// TIA Portal project "Project2" (V17)

(* hardware
DEVICE "S7-1500/ET200MP station_1"  S7-1500 station
   slot 0: "Rail_0"  Rack  6ES7 590-1***0-0AA0
   slot 1: "PLC_2"  CPU 1515-2 PN  6ES7 515-2AM00-0AB0  V1.8
      slot 3: "CPU display_1"  6ES7591-1BA00-0AA0
      slot 32768: "PROFINET interface_1"  X1
         slot 32769: "Port_1"  X1 P1
         slot 32770: "Port_2"  X1 P2
      slot 33024: "PROFINET interface_2"  X2
         slot 33025: "Port_1"  X2 P1
*)

// ===== PLC "PLC_2"  CPU 1515-2 PN =====

// folder: UDT/S2-Process Function Unit

TYPE "UDT_IS28xx_To_Plc"
   STRUCT
      iTriggerReady : Bool;   // This bit indicates when an In-Sight device can accept a new trigger via the Trigger bit. This field is true when the Trigger Enable bit is set, and the vision system is not currently acquiring an image.
      iTriggerAck : Bool;   // This bit indicates when an In-Sight device is successfully triggered via the Trigger bit. The Trigger Acknowledge bit stays set until the Trigger bit is cleared.
      iExposureComplete : Bool;   // This bit is set when the vision system image sensor is no longer exposed to light. It is used to indicate that the part being inspected can be moved from under the vision system's field of view.
      iAcquisitionError : Bool;   // This bit is set when an In-Sight device fails to acquire an image for one of the following reasons:
      iOfflineReason_1 : Bool;   // OfflineReason_1
      iOfflineReason_2 : Bool;   // OfflineReason_2
      iOfflineReason_3 : Bool;   // OfflineReason_3
      iSystemOnline : Bool;   // This bit indicates that the In-Sight device is online and the $System.OnlineEnabled tag is True.
      iReserve_1 : Byte;   // Reserve1
      iAcquisitonID : Int;   // This ID increments on the completion of every acquisition, regardless of the trigger source, and can be used to synchronize an acquisition with its Inspection Result. The Acquisition ID is changed on the start of an acquisition. If the PLC is the trigger source, the Acquisition ID is set prior to setting the Trigger Acknowledge bit.
      iReserve_2 : Bool;   // Reserve2
      iInspectionComplete : Bool;   // This bit is toggled upon the completion of an inspection.
      iResultBufferOverRun : Bool;   // This bit is set when the Enable Results Buffer bit is set, and there are more results than the result queue can hold.
      iResultValid : Bool;   // This bit is set when the Inspected Image ID, Inspection Result Code and Inspection Results fields are valid. The bit is cleared when the Inspection Results Acknowledge bit is set.
      iCommandExecuted : Bool;   // This bit is set while a command execution is in progress.
      iCommandComplete : Bool;   // This bit is set when the command execution is completed, and cleared when the Execute Command bit has been cleare
      iCommandFailed : Bool;   // This bit is set on the completion of a command, if the command has failed to execute successfully, or if an unknown Command ID was set.
      iSetUserDataAck : Bool;   // This bit is set to acknowledge completion of the Set User Data command.
      iJobPass : Bool;   // This bit indicates the pass and/or fail state of the inspection.
      iReserve_3 : Bool;   // Reserve3
      iReserve_4 : Bool;   // Reserve4
      iReserve_5 : Bool;   // Reserve5
      iReserve_6 : Bool;   // Reserve6
      iReserve_7 : Bool;   // Reserve7
      iReserve_8 : Bool;   // Reserve8
      iError : Bool;   // This bit is set when an error has occurred, which is defined in the Error ID field.
      iErrorID : Int;   // See Error ID codes.
      iCurrentRunningJobID : Int;   // These bits indicate the pre-added number of the current job filename. A job ID is a 16 bit number from 0 to 65535, but the PLC function can only load job IDs between 0‑999.
      iCommandResultCode : Int;   // This field is used to indicate the reason a command failed to execute successfully (the code is specific to the command executed):
      iExternalSoftEventAck : Byte;   // The External Event Acknowledge will be generated after the associated script finishes its execution
      iInspectionResultData : Struct
         iInspectionID : Int;   // The acquisition ID associated with this set of results.
         iInspectionResultCode : Int;   // These bytes are used to pass the user-defined result code. The inspection result code is defined by the Result Code parameter of the WriteResultsBuffer function
         iInspectionResult : Array[1..60] of Byte;   // These bytes of the inspection tool results can be written to the currently enabled factory communication protocol via the WriteResultsBuffer function.
      END_STRUCT;
   END_STRUCT;
END_TYPE

TYPE "UDT_Plc_To_IS28xx"
   STRUCT
      qTriggerEnable : Bool;   // This field is set to enable triggering via the Trigger bit. Clear this bit to disable the network triggering mechanism
      qTrigger : Bool;   // Setting the Trigger bit will trigger an acquisition on the vision system. The Trigger Enable bit must also be set
      qClearExposureComplete : Bool;   // When this signal is held high, the Exposure Complete status will remain reset. Once this signal is set to low, the Exposure Complete status will be set to high on the next exposure completion.
      qReserve_1 : Bool;   // Reserve_1
      qReserve_2 : Bool;   // Reserve_2
      qReserve_3 : Bool;   // Reserve_3
      qReserve_4 : Bool;   // Reserve_4
      qSetOffline : Bool;   // When this bit is set, the In-Sight vision system is paused and the state of the $System.OnlineEnabledComm is false
      qBufferResultEnable : Bool;   // When this bit is set, the Inspection ID, Inspection Result and Inspection Results fields are held constant until the Inspection Results Acknowledge field has acknowledged them and been set. Up to 16 sets of results are held in the buffer. Each result must be explicitly acknowledged using the Inspection Results Acknowledge signal.
      qInspectionResultAck : Bool;   // When the Buffer Results Enable bit is set, the Inspection Results Acknowledge bit acknowledges that the PLC has received the Inspected Image ID, Inspection Result Code and Inspection Results data.
      qSetUserData : Bool;   // This bit is used to signal that new User Data is available to be read in the vision system. After latching the entire User Data area into a holding buffer, the vision system will indicate to the PLC that it has read the data, and it can start loading new data into the buffer, if required, by issuing the Set User Data Acknowledge signal.
      qExecuteCommand : Bool;   // When the Execute Command bit is set to high, the Command ID signal is read by the vision system and the associated command is executed. The signal must be held high until the Command Completed bit is set. Once the Command Completed bit is set, clearing the Execute Command bit also clears the Command Completed bit.
      qReserve_5 : Bool;   // Reserve_5
      qReserve_6 : Bool;   // Reserve_6
      qReserve_7 : Bool;   // Reserve_7
      qClearError : Bool;   // When this bit is set, it clears the Error and Error ID signals; the Clear Error bit need to be held high until the Error bit is cleared. If an error is queued, clearing this bit causes the Error and Error ID signals to be set to the next queued error code.
      qCommandID : Int;   // This field indicates the command that will be executed on the rising edge of the Execute Command bit. This signal should not be changed until the Command Completed bit has been set.
      qSoftControlInput : Byte;   // Setting the External Event allows the PLC to trigger an associated event in the Spreadsheet.
      qUserData : Array[1..60] of Byte;   // Data buffer which can be read into the spreadsheet using the ReadUserDataBuffer function. The buffer is written exactly as it appears in the PLC
   END_STRUCT;
END_TYPE

// folder: (top level)

ORGANIZATION_BLOCK "Main"   // OB1, LAD, ProgramCycle
TITLE = "Main Program Sweep (Cycle)"
{ S7_Optimized_Access := 'TRUE' }
VERSION : 0.1
   VAR_INPUT
      Initial_Call : Bool;   // Initial call of this OB
      Remanence : Bool;   // =True, if remanent data are available
   END_VAR
   VAR_TEMP
      OB1_EV_CLASS : Byte;   // Bits 0-3 = 1 (Coming event), Bits 4-7 = 1 (Event class 1)
      OB1_SCAN_1 : Byte;   // 1 (Cold restart scan 1 of OB 1), 3 (Scan 2-n of OB 1)
      OB1_PRIORITY : Byte;   // Priority of OB Execution
      OB1_OB_NUMBR : Byte;   // 1 (Organization block 1, OB1)
      OB1_RESERVED_1 : Byte;   // Reserved for system
      OB1_RESERVED_2 : Byte;   // Reserved for system
      OB1_PREV_CYCLE : Int;   // Cycle time of previous OB1 scan (milliseconds)
      OB1_MIN_CYCLE : Int;   // Minimum cycle time of OB1 (milliseconds)
      OB1_MAX_CYCLE : Int;   // Maximum cycle time of OB1 (milliseconds)
      OB1_DATE_TIME : Date_And_Time;   // Date and time OB1 started
   END_VAR
BEGIN
END_ORGANIZATION_BLOCK

// ===== library types =====

// folder: S2-Process Function Unit

FUNCTION_BLOCK "PR_CognexISCamera_Profinet"   // FB365, LAD
TITLE = Cognex2D_4Feature / Cognex Camera Module
{ S7_Optimized_Access := 'TRUE' }
AUTHOR : Deepak.Jagtap
FAMILY : WIPROPARI
NAME : S21006022005
VERSION : 0.1
// |============================================================================|
// BLOCK:Cognex Camera Module
// Item Code : SMxxxxx
// Owner:Precision Automation & Robotics India Ltd.
// Author: DJ
// Release Date:04-04-2018
// Version:0.1
// V0.1-Initial release
// |============================================================================|
// Block Description: This block is used for interface of Cognex Camera via 
// profinet  and enter Job selection from outside the block.
// |============================================================================|
// Errors:
// qErrTriggerTimeOut: Trigger TimeOut Error Occured
// qErrAcquiringTimeout: Acquiring TimeOut Error Occured
// qErrTriggerEnableTimeout: Trigger Enable TimeOut Occured
// qErrJobSelection: Job selection Error
// qBothStartOn: Both Start are ON
// ============================================================================|
// Dependency:
// Map Vision Input and Output from External IO address. Byte should be matched as per the block
// |============================================================================|
   VAR_INPUT
      iResetFault : Bool;   // Reset Fault Input
      iAutorunning : Bool;   // Autorunning Input
      iStartJobSelection : Bool;   // start job selection / Start for Job Selection
      iStartInspection : Bool;   // Start for Inspection / start inspection
      iRetryCount : Int;   // Retry Count eg:3,4 etc / retry count
      iRetryPB : Bool;
      iJobID : Int;   // Enter Job ID / job id
      iTriggerEnableTimeoutTime : Time;   // Trigger Enable TimeOut Time Delay
      iTriggerTimeoutTime : Time;   // Trigger TimeOut Time Delay
      iAcquiringTimeOutTime : Time;   // Acquiring TimeOut Time Delay
   END_VAR
   VAR_OUTPUT
      qJobPass : Bool;   // Job Pass In Inspection
      qJobFail : Bool;   // Job Failed In Inspection
      qJobSelectionOver : Bool;   // Connect Job Selection over bit / job selection over
      qJobInspectionOver : Bool;   // Inspection Over Output
      qVisionOnline : Bool;   // Insight Vision Is In Online
      qVisionOfflineReason1 : Bool;   // Insight Vision Offline Due To: The vision system's job is being modified
      qVisionOfflineReason2 : Bool;   // Insight Vision Offline Due To: A discrete signal is holding the vision system Offline
      qVisionOfflineReason3 : Bool;   // Insight Vision Offline Due To: A communications protocol is holding the vision system Offline
      qErrBothStartOn : Bool;   // Both Start are On / both start on
      qErrJobSelection : Bool;   // Job selection Error Occur / error job selection
      qErrTriggerEnableTimeout : Bool;   // Trigger Enable TimeOut Error
      qErrTriggerTimeOut : Bool;   // Trigger TimeOut Error
      qErrAcquiringTimeOut : Bool;   // Acquiring TimeOut Error
   END_VAR
   VAR_IN_OUT
      iqInputAddrs : ANY;   // Input HW Address P#I120.0 BYTE 74
      iqOutputAddrs : ANY;   // Input HW Address P#Q120.0 BYTE 68
      iqRetryCount : Int;   // Retry Count Display / Retry count
      iqRunningJobID : Int;   // Running job ID
      iqInsight_Camera : Struct   // Insight Camera PZD
         Vision_Input : Struct
            "iTrigger Ready" : Bool;
            "iTrigger Ack" : Bool;
            iExposureComplete : Bool;
            "iMissed Ack" : Bool;
            "iOffline Reason_0" : Bool;
            "iOffline Reason_1" : Bool;
            "iOffline Reason_2" : Bool;
            iOnline : Bool;
            Acquisition_ID : Byte;
            Acquisition_ID_1 : Byte;
            iSystemBusy : Bool;
            "iInspection Completed" : Bool;
            "iResults Buffer Overrun" : Bool;
            "iResults Valid" : Bool;
            iCommandExecuting : Bool;
            iCommandComplete : Bool;
            "iCommand Failed" : Bool;
            iSetUserDataAck : Bool;
            iJobPass : Bool;
            iReserved : Bool;
            iReserved_1 : Bool;
            iReserved_2 : Bool;
            iReserved_3 : Bool;
            iReserved_4 : Bool;
            iReserved_5 : Bool;
            iError : Bool;
            iErrorCode : Int;
            iCommandControlInput : Int;
            SoftEventControlInput : Byte;
            iInspection_ID : Byte;
            iInspection_ID_1 : Byte;
            iInspection_ResultCode : Byte;
            iInspection_ResultCode_1 : Byte;
            iInspection_Result : Array[213..277] of Byte;
         END_STRUCT;
         Vision_Output : Struct
            "qTrigger Enable" : Bool;
            qTrigger : Bool;
            qClearExposureComplete : Bool;
            qReserved_1 : Bool;
            qReserved_2 : Bool;
            qReserved_3 : Bool;
            qReserved_4 : Bool;
            "qSet Offline" : Bool;
            "qBuffer Results Enable" : Bool;
            "qInspection Results Ack" : Bool;
            qSetUserData : Bool;
            qExecuteCommand : Bool;
            qReserved : Bool;
            qReserved_5 : Bool;
            qReserved_6 : Bool;
            qClearError : Bool;
            qCommandControl : Word;
            "Soft Event Control" : Byte;
            qUser_Data : Array[205..268] of Byte;
         END_STRUCT;
      END_STRUCT;
   END_VAR
   VAR
      sResetFaults : Bool;   // Reset Faults
      sInspectionComplete : Bool;   // Inspection Complete
      TriggerTimeout : TON_TIME;   // TriggerTimeout Timer
      TriggerEnableTimeout : TON_TIME;   // TriggerEnableTimeout Timer
      AcquiringTimeOut : TON_TIME;   // AcquiringTimeOut Timer
      ResultTimer : TON_TIME;   // ResultTimer
      sPulse : Array[0..11] of Bool;   // Array of Pulses
      sJobPass : Bool;   // Stat Bit of Job Pass
      sVisionInputCmdControlIP : Int;
      sJobFail : Bool;   // Stat Bit of Job Fail
      sJobLoadcompleted : Bool;
      sErrTriggerTimeOut : Bool;   // Error Trigger Time Out
      sErrJobSelection : Bool;
      sBothStartOn : Bool;
      sJobSelectionOver : Bool;
      sJobInspectionOver : Bool;
      sErrAcquiringTimeOut : Bool;   // Error Acquiring Time Out
      sErrTriggerEnableTimeout : Bool;   // Error Trigger Enable Time Out
      sVisionOutput_Trigger : Bool;   // Vision Outpur Trigger
      sRetryCountOver : Bool;
      sInitialPulse : Bool;
      sProgramEcho : TON_TIME;
      sExposureTimerStar1 : Bool;
      sExposureTimerStart : Bool;
      sExposureTimer : TON_TIME;
      sExecDelayTimer : TON_TIME;
      sRetry : TON_TIME;
   END_VAR
   VAR_TEMP
      tInspectionID : Int;
      tResultCode : Int;
   END_VAR
   VAR_TEMP   // added for the SCL form of the ladder/FBD networks
      _w1 : Bool;
      _w2 : Bool;
      _w3 : Bool;
      _w4 : Bool;
   END_VAR
BEGIN

REGION Network 1: Header
   // ==============================================================================
   //  Company: Precision Automation & Robotics India Ltd. 
   // ------------------------------------------------------------------------------
   //  Item Code: S21006022005
   //  Author/Created by: Deepak.Jagtap
   //  Reviewed/Checked by: Atul P
   //  First Release on: 04-04-2018
   //  Latest update on:
   // ------------------------------------------------------------------------------
   //  Tested with: CPU firmware, model or simulator testing
   //  Engineering/Editor: TIA Portal V15.1
   // ------------------------------------------------------------------------------
   //  Restrictions:
   //  Dependencies/Requirements:
   // iqInsight_Camera	Struct
   // Map Vision Input and Output from with External IO address
   // ------------------------------------------------------------------------------
   //  Change Log:
   //  Ver.	Date		Changed by		Details of changes
   //  1.0	04-04-2018	Deepak.Jagtap            	First release version
   // 
   // ------------------------------------------------------------------------------
   //  Functionality: This block is used for interface of Cognex Camera via 
   // profinet.
   // 
   //  Inputs
   // iResetFault	Bool
   // iAutorunning	Bool
   // iStartJobSelection	Bool
   // iStartInspection	Bool
   // iRetryCount	Int
   // iJobID	Int
   // iTriggerEnableTimeoutTime	Time
   // iTriggerTimeoutTime	Time
   // iAcquiringTimeOutTime	Time
   // 
   //  Outputs
   // qJobPass	Bool
   // qJobFail	Bool
   // qJobSelectionOver	Bool
   // qJobInspectionOver	Bool
   // qVisionOnline	Bool
   // qVisionOfflineReason1	Bool
   // qVisionOfflineReason2	Bool
   // qVisionOfflineReason3	Bool
   // qErrBothStartOn	Bool
   // qErrJobSelection	Bool
   // qErrTriggerEnableTimeout	Bool
   // qErrTriggerTimeOut	Bool
   // qErrAcquiringTimeOut	Bool
   // 
   //  In-outs
   // iqInputAddrs	Any
   // iqOutputAddrs	Any
   // iqRetryCount	Int
   // iqRunningJobID	Int
   // iqInsight_Camera	Struct
   // 
   // ------------------------------------------------------------------------------
   //  Errors reported:
   //  1.qErrTriggerTimeOut : Error trigger timeout
   // 2. qErrAcquiringTimeOut;Acquiring Time Out
   // 3. qErrTriggerEnableTimeout:Trigger Enable Time Out
   // 4. qErrBothStartOn:both start on
   // 5. qErrJobSelection:error job selection
   //  Messages reported:
   //  1. Message 1 present
   //  2. Message 2 present
   // ==============================================================================
END_REGION

REGION Network 2: Read Data From Input Area
   // Read Data From Input Area
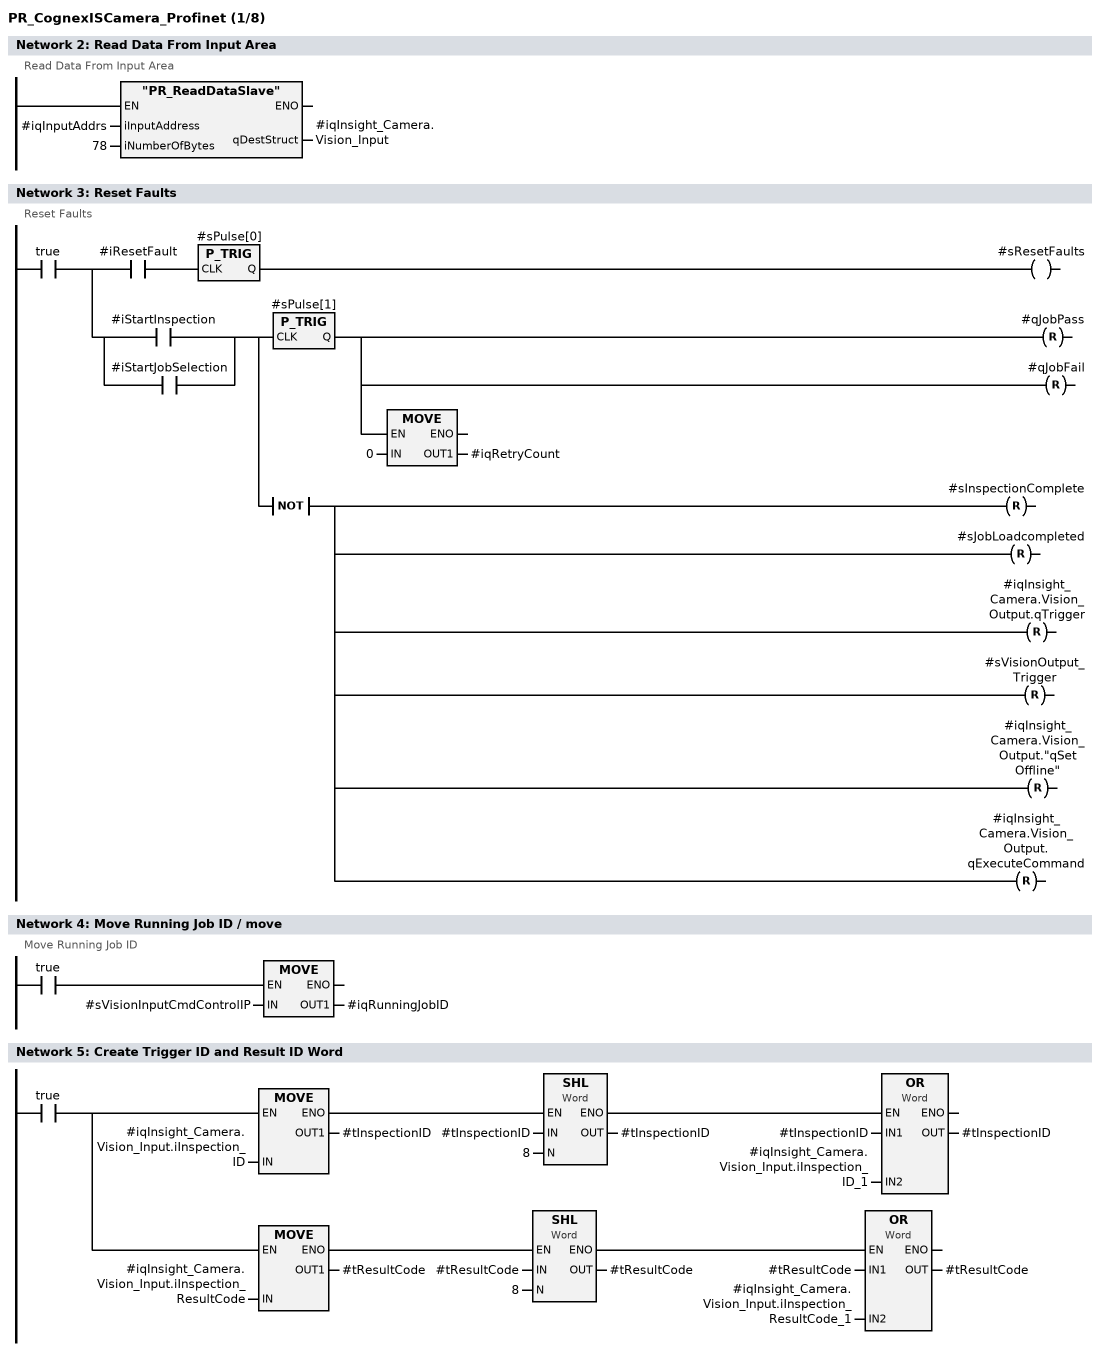
   RUNG wire#powerrail
      "PR_ReadDataSlave"(iInputAddress := #iqInputAddrs, iNumberOfBytes := 78, qDestStruct => #iqInsight_Camera.Vision_Input)
   END_RUNG
   // the same network as SCL:
   "PR_ReadDataSlave"(iInputAddress := #iqInputAddrs,
                      iNumberOfBytes := 78,
                      qDestStruct => #iqInsight_Camera.Vision_Input);
END_REGION

REGION Network 3: Reset Faults
   // Reset Faults
   RUNG wire#powerrail
      Contact( true )
      wire#w1
      Contact( #iResetFault )
      P_Trig( #sPulse[0] )
      Coil( #sResetFaults )
   END_RUNG
   RUNG wire#w1
      Contact( #iStartInspection )
      wire#w2
      P_Trig( #sPulse[1] )
      wire#w3
      R_Coil( #qJobPass )
   END_RUNG
   RUNG wire#w1
      Contact( #iStartJobSelection )
   END_RUNG wire#w2
   RUNG wire#w3
      R_Coil( #qJobFail )
   END_RUNG
   RUNG wire#w3
      Move(in := 0, out1 => #iqRetryCount)
   END_RUNG
   RUNG wire#w2
      Not()
      wire#w4
      R_Coil( #sInspectionComplete )
   END_RUNG
   RUNG wire#w4
      R_Coil( #sJobLoadcompleted )
   END_RUNG
   RUNG wire#w4
      R_Coil( #iqInsight_Camera.Vision_Output.qTrigger )
   END_RUNG
   RUNG wire#w4
      R_Coil( #sVisionOutput_Trigger )
   END_RUNG
   RUNG wire#w4
      R_Coil( #iqInsight_Camera.Vision_Output."qSet Offline" )
   END_RUNG
   RUNG wire#w4
      R_Coil( #iqInsight_Camera.Vision_Output.qExecuteCommand )
   END_RUNG
   // the same network as SCL:
   #_w1 := true AND #iResetFault;
   #_w2 := #_w1 AND NOT #sPulse[0];   // rising edge
   #sPulse[0] := #_w1;
   #sResetFaults := #_w2;
   #_w3 := true AND (#iStartInspection OR #iStartJobSelection);
   #_w4 := #_w3 AND NOT #sPulse[1];   // rising edge
   #sPulse[1] := #_w3;
   IF #_w4 THEN
       #qJobPass := FALSE;
       #qJobFail := FALSE;
       #iqRetryCount := 0;
   END_IF;
   IF NOT #_w3 THEN
       #sInspectionComplete := FALSE;
       #sJobLoadcompleted := FALSE;
       #iqInsight_Camera.Vision_Output.qTrigger := FALSE;
       #sVisionOutput_Trigger := FALSE;
       #iqInsight_Camera.Vision_Output."qSet Offline" := FALSE;
       #iqInsight_Camera.Vision_Output.qExecuteCommand := FALSE;
   END_IF;
END_REGION

REGION Network 4: Move Running Job ID / move
   // Move Running Job ID
   RUNG wire#powerrail
      Contact( true )
      Move(in := #sVisionInputCmdControlIP, out1 => #iqRunningJobID)
   END_RUNG
   // the same network as SCL:
   IF true THEN #iqRunningJobID := #sVisionInputCmdControlIP; END_IF;
END_REGION

REGION Network 5: Create Trigger ID and Result ID Word
   IF true THEN
       #tInspectionID := #iqInsight_Camera.Vision_Input.iInspection_ID;
       #tInspectionID := SHL(IN := #tInspectionID, N := 8);
       #tInspectionID := #tInspectionID OR #iqInsight_Camera.Vision_Input.iInspection_ID_1;
       #tResultCode := #iqInsight_Camera.Vision_Input.iInspection_ResultCode;
       #tResultCode := SHL(IN := #tResultCode, N := 8);
       #tResultCode := #tResultCode OR #iqInsight_Camera.Vision_Input.iInspection_ResultCode_1;
   END_IF;
END_REGION

REGION Network 6: Trigger Enable through Job Selection / Camera Trigger Enable
   // Trigger Enable through Job Selection
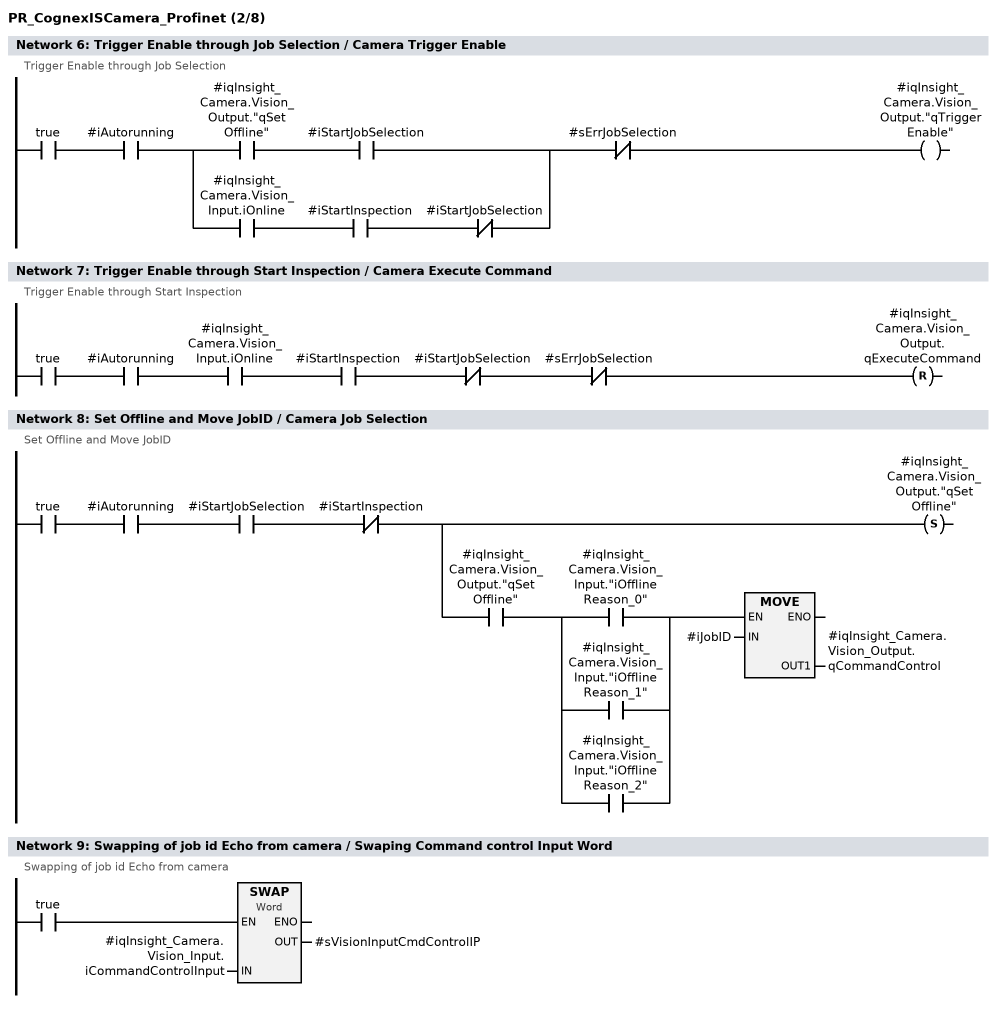
   RUNG wire#powerrail
      Contact( true )
      Contact( #iAutorunning )
      wire#w1
      Contact( #iqInsight_Camera.Vision_Output."qSet Offline" )
      Contact( #iStartJobSelection )
      wire#w2
      I_Contact( #sErrJobSelection )
      Coil( #iqInsight_Camera.Vision_Output."qTrigger Enable" )
   END_RUNG
   RUNG wire#w1
      Contact( #iqInsight_Camera.Vision_Input.iOnline )
      Contact( #iStartInspection )
      I_Contact( #iStartJobSelection )
   END_RUNG wire#w2
   // the same network as SCL:
   #iqInsight_Camera.Vision_Output."qTrigger Enable" := true AND #iAutorunning AND ((#iqInsight_Camera.Vision_Output."qSet Offline" AND #iStartJobSelection) OR (#iqInsight_Camera.Vision_Input.iOnline AND #iStartInspection AND NOT #iStartJobSelection)) AND NOT #sErrJobSelection;
END_REGION

REGION Network 7: Trigger Enable through Start Inspection / Camera Execute Command
   // Trigger Enable through Start Inspection
   RUNG wire#powerrail
      Contact( true )
      Contact( #iAutorunning )
      Contact( #iqInsight_Camera.Vision_Input.iOnline )
      Contact( #iStartInspection )
      I_Contact( #iStartJobSelection )
      I_Contact( #sErrJobSelection )
      R_Coil( #iqInsight_Camera.Vision_Output.qExecuteCommand )
   END_RUNG
   // the same network as SCL:
   IF true AND #iAutorunning AND #iqInsight_Camera.Vision_Input.iOnline AND #iStartInspection AND NOT #iStartJobSelection AND NOT #sErrJobSelection THEN
       #iqInsight_Camera.Vision_Output.qExecuteCommand := FALSE;
   END_IF;
END_REGION

REGION Network 8: Set Offline and Move JobID / Camera Job Selection
   // Set Offline and Move JobID
   RUNG wire#powerrail
      Contact( true )
      Contact( #iAutorunning )
      Contact( #iStartJobSelection )
      I_Contact( #iStartInspection )
      wire#w1
      S_Coil( #iqInsight_Camera.Vision_Output."qSet Offline" )
   END_RUNG
   RUNG wire#w1
      Contact( #iqInsight_Camera.Vision_Output."qSet Offline" )
      wire#w2
      Contact( #iqInsight_Camera.Vision_Input."iOffline Reason_0" )
      wire#w3
      Move(in := #iJobID, out1 => #iqInsight_Camera.Vision_Output.qCommandControl)
   END_RUNG
   RUNG wire#w2
      Contact( #iqInsight_Camera.Vision_Input."iOffline Reason_1" )
   END_RUNG wire#w3
   RUNG wire#w2
      Contact( #iqInsight_Camera.Vision_Input."iOffline Reason_2" )
   END_RUNG wire#w3
   // the same network as SCL:
   #_w1 := true AND #iAutorunning AND #iStartJobSelection AND NOT #iStartInspection;
   IF #_w1 THEN #iqInsight_Camera.Vision_Output."qSet Offline" := TRUE; END_IF;
   IF #_w1 AND #iqInsight_Camera.Vision_Output."qSet Offline" AND (#iqInsight_Camera.Vision_Input."iOffline Reason_0" OR #iqInsight_Camera.Vision_Input."iOffline Reason_1" OR #iqInsight_Camera.Vision_Input."iOffline Reason_2") THEN
       #iqInsight_Camera.Vision_Output.qCommandControl := #iJobID;
   END_IF;
END_REGION

REGION Network 9: Swapping of job id Echo from camera / Swaping Command control Input Word
   // Swapping of job id Echo from camera
   IF true THEN
       #sVisionInputCmdControlIP := SWAP(#iqInsight_Camera.Vision_Input.iCommandControlInput);
   END_IF;
END_REGION

REGION Network 10: Initiate Job Load / Camera Execute Command
   // Initiate Job Load
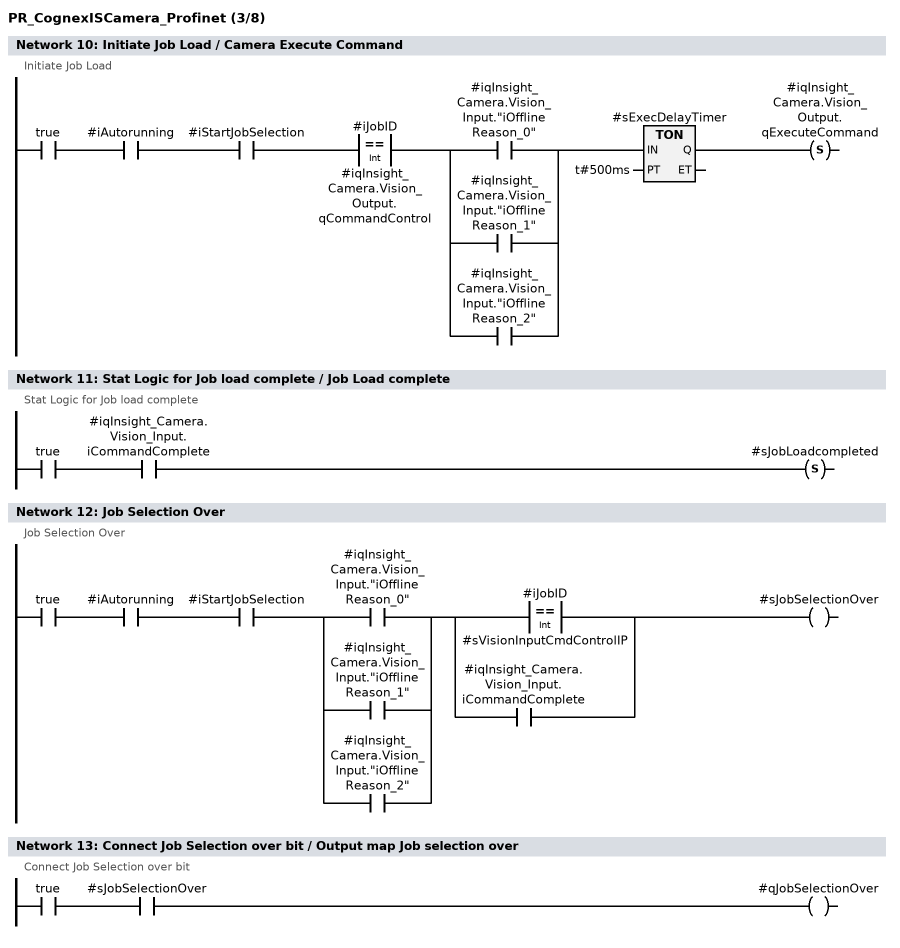
   #sExecDelayTimer(IN := true AND #iAutorunning AND #iStartJobSelection AND (#iJobID = #iqInsight_Camera.Vision_Output.qCommandControl) AND (#iqInsight_Camera.Vision_Input."iOffline Reason_0" OR #iqInsight_Camera.Vision_Input."iOffline Reason_1" OR #iqInsight_Camera.Vision_Input."iOffline Reason_2"),   // TON
                    PT := t#500ms);
   IF #sExecDelayTimer.Q THEN #iqInsight_Camera.Vision_Output.qExecuteCommand := TRUE; END_IF;
END_REGION

REGION Network 11: Stat Logic for Job load complete / Job Load complete
   // Stat Logic for Job load complete
   RUNG wire#powerrail
      Contact( true )
      Contact( #iqInsight_Camera.Vision_Input.iCommandComplete )
      S_Coil( #sJobLoadcompleted )
   END_RUNG
   // the same network as SCL:
   IF true AND #iqInsight_Camera.Vision_Input.iCommandComplete THEN #sJobLoadcompleted := TRUE; END_IF;
END_REGION

REGION Network 12: Job Selection Over
   // Job Selection Over
   RUNG wire#powerrail
      Contact( true )
      Contact( #iAutorunning )
      Contact( #iStartJobSelection )
      wire#w1
      Contact( #iqInsight_Camera.Vision_Input."iOffline Reason_0" )
      wire#w2
      { S7_Templates := "SrcType := Int" } EQ_Contact(in1 := #iJobID, in2 := #sVisionInputCmdControlIP)
      wire#w3
      Coil( #sJobSelectionOver )
   END_RUNG
   RUNG wire#w1
      Contact( #iqInsight_Camera.Vision_Input."iOffline Reason_1" )
   END_RUNG wire#w2
   RUNG wire#w1
      Contact( #iqInsight_Camera.Vision_Input."iOffline Reason_2" )
   END_RUNG wire#w2
   RUNG wire#w2
      Contact( #iqInsight_Camera.Vision_Input.iCommandComplete )
   END_RUNG wire#w3
   // the same network as SCL:
   #sJobSelectionOver := true AND #iAutorunning AND #iStartJobSelection AND (#iqInsight_Camera.Vision_Input."iOffline Reason_0" OR #iqInsight_Camera.Vision_Input."iOffline Reason_1" OR #iqInsight_Camera.Vision_Input."iOffline Reason_2") AND ((#iJobID = #sVisionInputCmdControlIP) OR #iqInsight_Camera.Vision_Input.iCommandComplete);
END_REGION

REGION Network 13: Connect Job Selection over bit / Output map Job selection over
   // Connect Job Selection over bit
   RUNG wire#powerrail
      Contact( true )
      Contact( #sJobSelectionOver )
      Coil( #qJobSelectionOver )
   END_RUNG
   // the same network as SCL:
   #qJobSelectionOver := true AND #sJobSelectionOver;
END_REGION

REGION Network 14: Reset Offline / Camera Job Selection reset
   // Reset Offline / "#iqInsight_Camera.Vision_Output.qSet Offline" and "#iqInsight_Camera.Vision_Output.qExecuteCommand"  Reset coil removed while block comparision
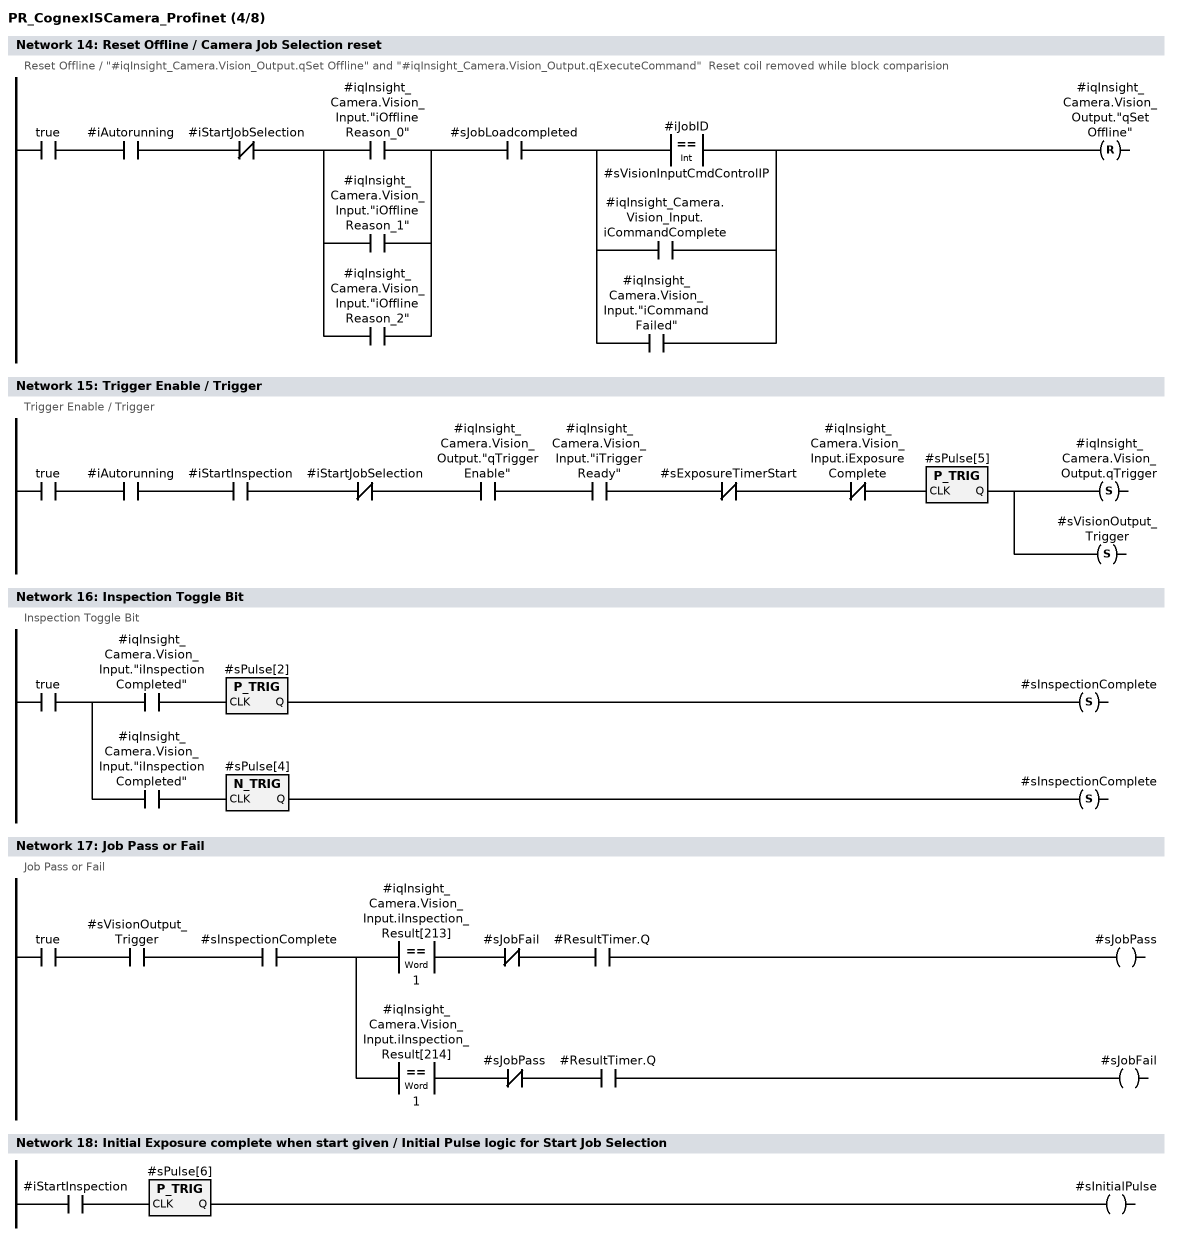
   RUNG wire#powerrail
      Contact( true )
      Contact( #iAutorunning )
      I_Contact( #iStartJobSelection )
      wire#w1
      Contact( #iqInsight_Camera.Vision_Input."iOffline Reason_0" )
      wire#w2
      Contact( #sJobLoadcompleted )
      wire#w3
      { S7_Templates := "SrcType := Int" } EQ_Contact(in1 := #iJobID, in2 := #sVisionInputCmdControlIP)
      wire#w4
      R_Coil( #iqInsight_Camera.Vision_Output."qSet Offline" )
   END_RUNG
   RUNG wire#w1
      Contact( #iqInsight_Camera.Vision_Input."iOffline Reason_1" )
   END_RUNG wire#w2
   RUNG wire#w1
      Contact( #iqInsight_Camera.Vision_Input."iOffline Reason_2" )
   END_RUNG wire#w2
   RUNG wire#w3
      Contact( #iqInsight_Camera.Vision_Input.iCommandComplete )
   END_RUNG wire#w4
   RUNG wire#w3
      Contact( #iqInsight_Camera.Vision_Input."iCommand Failed" )
   END_RUNG wire#w4
   // the same network as SCL:
   IF true AND #iAutorunning AND NOT #iStartJobSelection AND (#iqInsight_Camera.Vision_Input."iOffline Reason_0" OR #iqInsight_Camera.Vision_Input."iOffline Reason_1" OR #iqInsight_Camera.Vision_Input."iOffline Reason_2") AND #sJobLoadcompleted AND ((#iJobID = #sVisionInputCmdControlIP) OR #iqInsight_Camera.Vision_Input.iCommandComplete OR #iqInsight_Camera.Vision_Input."iCommand Failed") THEN
       #iqInsight_Camera.Vision_Output."qSet Offline" := FALSE;
   END_IF;
END_REGION

REGION Network 15: Trigger Enable / Trigger
   // Trigger Enable / Trigger
   RUNG wire#powerrail
      Contact( true )
      Contact( #iAutorunning )
      Contact( #iStartInspection )
      I_Contact( #iStartJobSelection )
      Contact( #iqInsight_Camera.Vision_Output."qTrigger Enable" )
      Contact( #iqInsight_Camera.Vision_Input."iTrigger Ready" )
      I_Contact( #sExposureTimerStart )
      I_Contact( #iqInsight_Camera.Vision_Input.iExposureComplete )
      P_Trig( #sPulse[5] )
      wire#w1
      S_Coil( #iqInsight_Camera.Vision_Output.qTrigger )
   END_RUNG
   RUNG wire#w1
      S_Coil( #sVisionOutput_Trigger )
   END_RUNG
   // the same network as SCL:
   #_w1 := true AND #iAutorunning AND #iStartInspection AND NOT #iStartJobSelection AND #iqInsight_Camera.Vision_Output."qTrigger Enable" AND #iqInsight_Camera.Vision_Input."iTrigger Ready" AND NOT #sExposureTimerStart AND NOT #iqInsight_Camera.Vision_Input.iExposureComplete;
   #_w2 := #_w1 AND NOT #sPulse[5];   // rising edge
   #sPulse[5] := #_w1;
   IF #_w2 THEN
       #iqInsight_Camera.Vision_Output.qTrigger := TRUE;
       #sVisionOutput_Trigger := TRUE;
   END_IF;
END_REGION

REGION Network 16: Inspection Toggle Bit
   // Inspection Toggle Bit
   RUNG wire#powerrail
      Contact( true )
      wire#w1
      Contact( #iqInsight_Camera.Vision_Input."iInspection Completed" )
      P_Trig( #sPulse[2] )
      S_Coil( #sInspectionComplete )
   END_RUNG
   RUNG wire#w1
      Contact( #iqInsight_Camera.Vision_Input."iInspection Completed" )
      N_Trig( #sPulse[4] )
      S_Coil( #sInspectionComplete )
   END_RUNG
   // the same network as SCL:
   #_w1 := true AND #iqInsight_Camera.Vision_Input."iInspection Completed";
   #_w2 := #_w1 AND NOT #sPulse[2];   // rising edge
   #sPulse[2] := #_w1;
   IF #_w2 THEN #sInspectionComplete := TRUE; END_IF;
   #_w3 := true AND #iqInsight_Camera.Vision_Input."iInspection Completed";
   #_w4 := NOT #_w3 AND #sPulse[4];   // falling edge
   #sPulse[4] := #_w3;
   IF #_w4 THEN #sInspectionComplete := TRUE; END_IF;
END_REGION

REGION Network 17: Job Pass or Fail
   // Job Pass or Fail
   RUNG wire#powerrail
      Contact( true )
      Contact( #sVisionOutput_Trigger )
      Contact( #sInspectionComplete )
      wire#w1
      { S7_Templates := "SrcType := Word" } EQ_Contact(in1 := #iqInsight_Camera.Vision_Input.iInspection_Result[213], in2 := 1)
      I_Contact( #sJobFail )
      Contact( #ResultTimer.Q )
      Coil( #sJobPass )
   END_RUNG
   RUNG wire#w1
      { S7_Templates := "SrcType := Word" } EQ_Contact(in1 := #iqInsight_Camera.Vision_Input.iInspection_Result[214], in2 := 1)
      I_Contact( #sJobPass )
      Contact( #ResultTimer.Q )
      Coil( #sJobFail )
   END_RUNG
   // the same network as SCL:
   #_w1 := true AND #sVisionOutput_Trigger AND #sInspectionComplete;
   #sJobPass := #_w1 AND (#iqInsight_Camera.Vision_Input.iInspection_Result[213] = 1) AND NOT #sJobFail AND #ResultTimer.Q;
   #sJobFail := #_w1 AND (#iqInsight_Camera.Vision_Input.iInspection_Result[214] = 1) AND NOT #sJobPass AND #ResultTimer.Q;
END_REGION

REGION Network 18: Initial Exposure complete when start given / Initial Pulse logic for Start Job Selection
   RUNG wire#powerrail
      Contact( #iStartInspection )
      P_Trig( #sPulse[6] )
      Coil( #sInitialPulse )
   END_RUNG
   // the same network as SCL:
   #_w1 := #iStartInspection AND NOT #sPulse[6];   // rising edge
   #sPulse[6] := #iStartInspection;
   #sInitialPulse := #_w1;
END_REGION

REGION Network 19: Exposure Timer 1
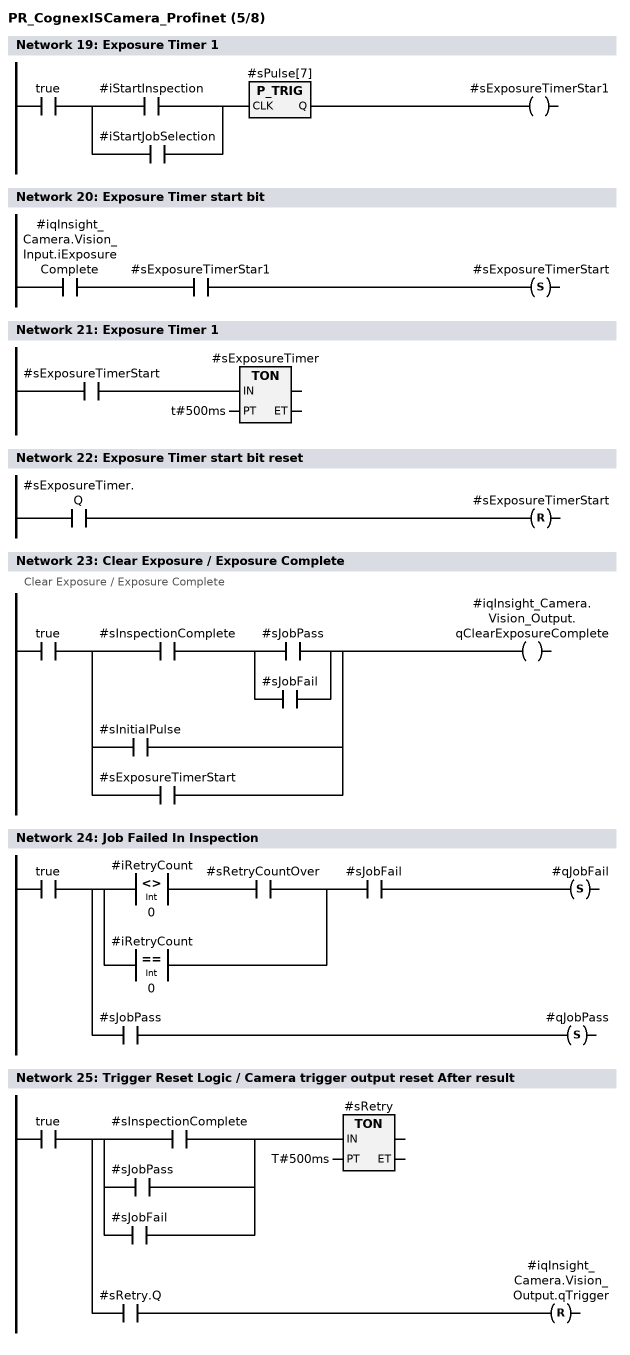
   RUNG wire#powerrail
      Contact( true )
      wire#w1
      Contact( #iStartInspection )
      wire#w2
      P_Trig( #sPulse[7] )
      Coil( #sExposureTimerStar1 )
   END_RUNG
   RUNG wire#w1
      Contact( #iStartJobSelection )
   END_RUNG wire#w2
   // the same network as SCL:
   #_w1 := true AND (#iStartInspection OR #iStartJobSelection);
   #_w2 := #_w1 AND NOT #sPulse[7];   // rising edge
   #sPulse[7] := #_w1;
   #sExposureTimerStar1 := #_w2;
END_REGION

REGION Network 20: Exposure Timer start bit
   RUNG wire#powerrail
      Contact( #iqInsight_Camera.Vision_Input.iExposureComplete )
      Contact( #sExposureTimerStar1 )
      S_Coil( #sExposureTimerStart )
   END_RUNG
   // the same network as SCL:
   IF #iqInsight_Camera.Vision_Input.iExposureComplete AND #sExposureTimerStar1 THEN
       #sExposureTimerStart := TRUE;
   END_IF;
END_REGION

REGION Network 21: Exposure Timer 1
   #sExposureTimer(IN := #sExposureTimerStart, PT := t#500ms);   // TON
END_REGION

REGION Network 22: Exposure Timer start bit reset
   RUNG wire#powerrail
      Contact( #sExposureTimer.Q )
      R_Coil( #sExposureTimerStart )
   END_RUNG
   // the same network as SCL:
   IF #sExposureTimer.Q THEN #sExposureTimerStart := FALSE; END_IF;
END_REGION

REGION Network 23: Clear Exposure / Exposure Complete
   // Clear Exposure / Exposure Complete
   RUNG wire#powerrail
      Contact( true )
      wire#w1
      Contact( #sInspectionComplete )
      wire#w2
      Contact( #sJobPass )
      wire#w3
      Coil( #iqInsight_Camera.Vision_Output.qClearExposureComplete )
   END_RUNG
   RUNG wire#w2
      Contact( #sJobFail )
   END_RUNG wire#w3
   RUNG wire#w1
      Contact( #sInitialPulse )
   END_RUNG wire#w3
   RUNG wire#w1
      Contact( #sExposureTimerStart )
   END_RUNG wire#w3
   // the same network as SCL:
   #iqInsight_Camera.Vision_Output.qClearExposureComplete := true AND ((#sInspectionComplete AND (#sJobPass OR #sJobFail)) OR #sInitialPulse OR #sExposureTimerStart);
END_REGION

REGION Network 24: Job Failed In Inspection
   RUNG wire#powerrail
      Contact( true )
      wire#w1
      { S7_Templates := "SrcType := Int" } NE_Contact(in1 := #iRetryCount, in2 := 0)
      Contact( #sRetryCountOver )
      wire#w2
      Contact( #sJobFail )
      S_Coil( #qJobFail )
   END_RUNG
   RUNG wire#w1
      { S7_Templates := "SrcType := Int" } EQ_Contact(in1 := #iRetryCount, in2 := 0)
   END_RUNG wire#w2
   RUNG wire#w1
      Contact( #sJobPass )
      S_Coil( #qJobPass )
   END_RUNG
   // the same network as SCL:
   IF true AND (((#iRetryCount <> 0) AND #sRetryCountOver) OR (#iRetryCount = 0)) AND #sJobFail THEN
       #qJobFail := TRUE;
   END_IF;
   IF true AND #sJobPass THEN #qJobPass := TRUE; END_IF;
END_REGION

REGION Network 25: Trigger Reset Logic / Camera trigger output reset After result
   #sRetry(IN := true AND (#sInspectionComplete OR #sJobPass OR #sJobFail), PT := T#500ms);   // TON
   IF true AND #sRetry.Q THEN #iqInsight_Camera.Vision_Output.qTrigger := FALSE; END_IF;
END_REGION

REGION Network 26: Retry Count Logic / CameraTrigger Enable on for retry count
   // Retry Count Logic
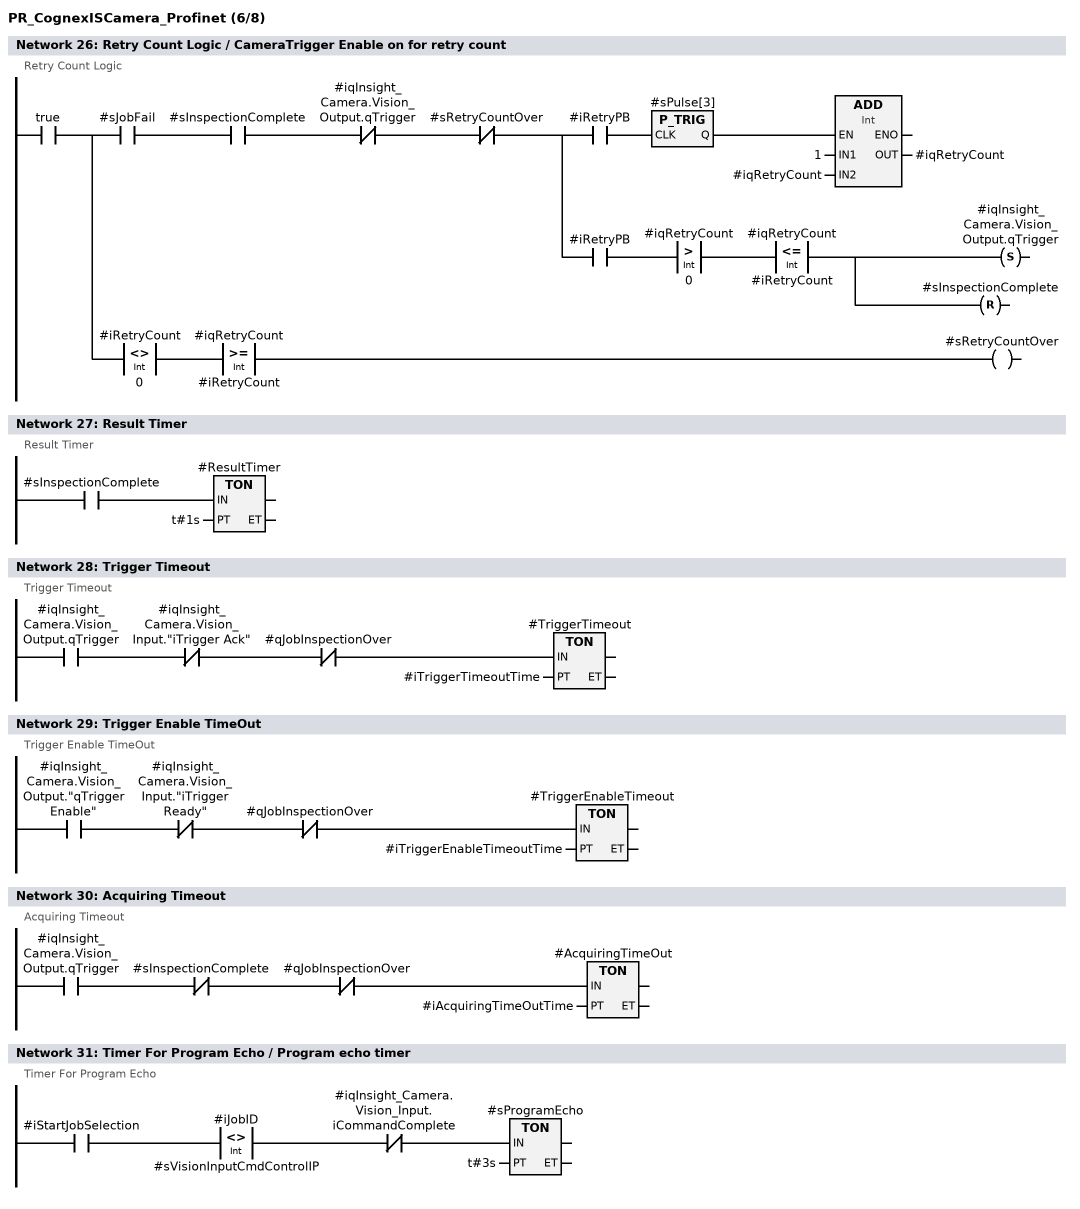
   RUNG wire#powerrail
      Contact( true )
      wire#w1
      Contact( #sJobFail )
      Contact( #sInspectionComplete )
      I_Contact( #iqInsight_Camera.Vision_Output.qTrigger )
      I_Contact( #sRetryCountOver )
      wire#w2
      Contact( #iRetryPB )
      P_Trig( #sPulse[3] )
      { S7_Templates := "SrcType := Int" } Add(in1 := 1, in2 := #iqRetryCount, out => #iqRetryCount)
   END_RUNG
   RUNG wire#w2
      Contact( #iRetryPB )
      { S7_Templates := "SrcType := Int" } GT_Contact(in1 := #iqRetryCount, in2 := 0)
      { S7_Templates := "SrcType := Int" } LE_Contact(in1 := #iqRetryCount, in2 := #iRetryCount)
      wire#w3
      S_Coil( #iqInsight_Camera.Vision_Output.qTrigger )
   END_RUNG
   RUNG wire#w3
      R_Coil( #sInspectionComplete )
   END_RUNG
   RUNG wire#w1
      { S7_Templates := "SrcType := Int" } NE_Contact(in1 := #iRetryCount, in2 := 0)
      { S7_Templates := "SrcType := Int" } GE_Contact(in1 := #iqRetryCount, in2 := #iRetryCount)
      Coil( #sRetryCountOver )
   END_RUNG
   // the same network as SCL:
   #_w1 := true AND #sJobFail AND #sInspectionComplete AND NOT #iqInsight_Camera.Vision_Output.qTrigger AND NOT #sRetryCountOver;
   #_w2 := #_w1 AND #iRetryPB;
   #_w3 := #_w2 AND NOT #sPulse[3];   // rising edge
   #sPulse[3] := #_w2;
   IF #_w3 THEN #iqRetryCount := 1 + #iqRetryCount; END_IF;
   IF #_w1 AND #iRetryPB AND (#iqRetryCount > 0) AND (#iqRetryCount <= #iRetryCount) THEN
       #iqInsight_Camera.Vision_Output.qTrigger := TRUE;
       #sInspectionComplete := FALSE;
   END_IF;
   #sRetryCountOver := true AND (#iRetryCount <> 0) AND (#iqRetryCount >= #iRetryCount);
END_REGION

REGION Network 27: Result Timer
   // Result Timer
   #ResultTimer(IN := #sInspectionComplete, PT := t#1s);   // TON
END_REGION

REGION Network 28: Trigger Timeout
   // Trigger Timeout
   #TriggerTimeout(IN := #iqInsight_Camera.Vision_Output.qTrigger AND NOT #iqInsight_Camera.Vision_Input."iTrigger Ack" AND NOT #qJobInspectionOver,   // TON
                   PT := #iTriggerTimeoutTime);
END_REGION

REGION Network 29: Trigger Enable TimeOut
   // Trigger Enable TimeOut
   #TriggerEnableTimeout(IN := #iqInsight_Camera.Vision_Output."qTrigger Enable" AND NOT #iqInsight_Camera.Vision_Input."iTrigger Ready" AND NOT #qJobInspectionOver,   // TON
                         PT := #iTriggerEnableTimeoutTime);
END_REGION

REGION Network 30: Acquiring Timeout
   // Acquiring Timeout
   #AcquiringTimeOut(IN := #iqInsight_Camera.Vision_Output.qTrigger AND NOT #sInspectionComplete AND NOT #qJobInspectionOver,   // TON
                     PT := #iAcquiringTimeOutTime);
END_REGION

REGION Network 31: Timer For Program Echo / Program echo timer
   // Timer For Program Echo
   #sProgramEcho(IN := #iStartJobSelection AND (#iJobID <> #sVisionInputCmdControlIP) AND NOT #iqInsight_Camera.Vision_Input.iCommandComplete,   // TON
                 PT := t#3s);
END_REGION

REGION Network 32: OutPuts
   // OutPuts
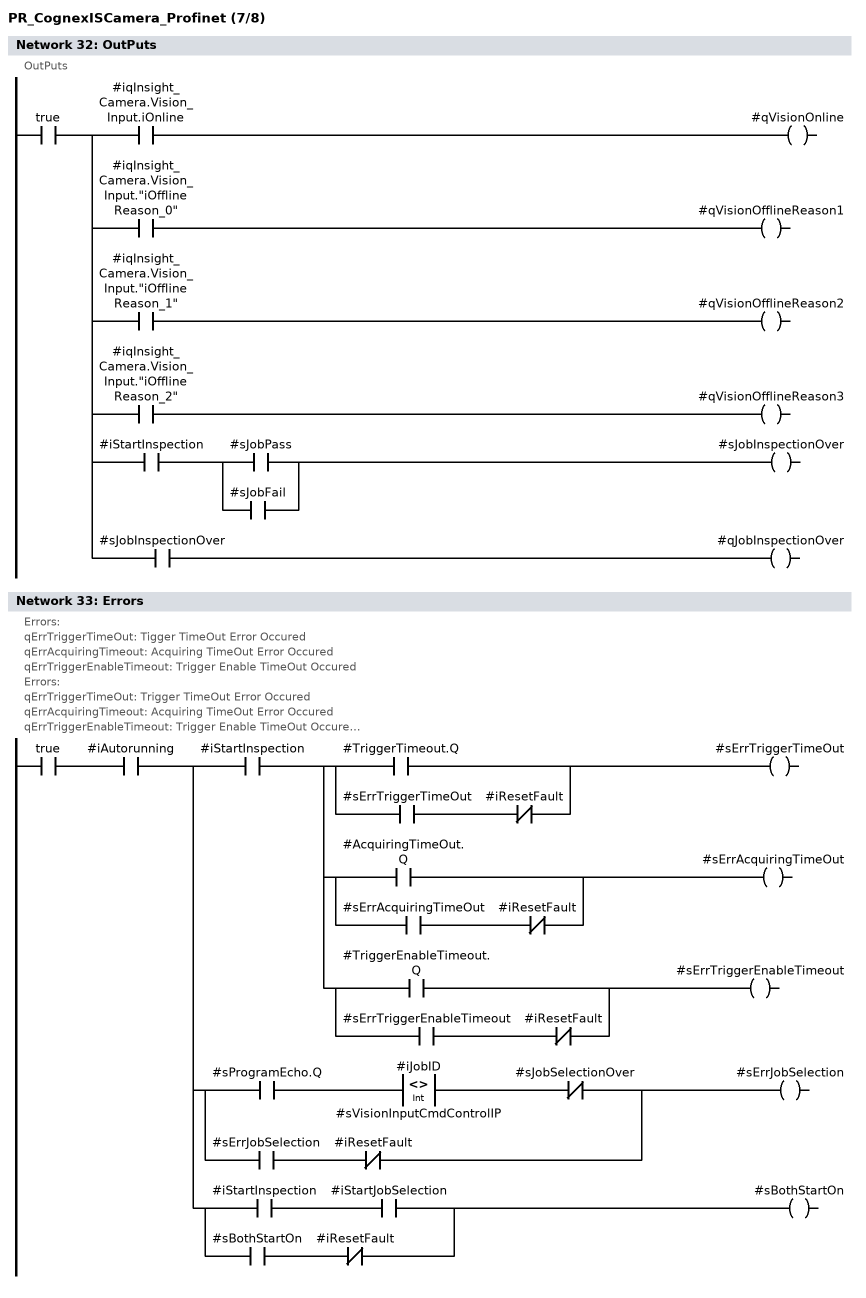
   RUNG wire#powerrail
      Contact( true )
      wire#w1
      Contact( #iqInsight_Camera.Vision_Input.iOnline )
      Coil( #qVisionOnline )
   END_RUNG
   RUNG wire#w1
      Contact( #iqInsight_Camera.Vision_Input."iOffline Reason_0" )
      Coil( #qVisionOfflineReason1 )
   END_RUNG
   RUNG wire#w1
      Contact( #iqInsight_Camera.Vision_Input."iOffline Reason_1" )
      Coil( #qVisionOfflineReason2 )
   END_RUNG
   RUNG wire#w1
      Contact( #iqInsight_Camera.Vision_Input."iOffline Reason_2" )
      Coil( #qVisionOfflineReason3 )
   END_RUNG
   RUNG wire#w1
      Contact( #iStartInspection )
      wire#w2
      Contact( #sJobPass )
      wire#w3
      Coil( #sJobInspectionOver )
   END_RUNG
   RUNG wire#w2
      Contact( #sJobFail )
   END_RUNG wire#w3
   RUNG wire#w1
      Contact( #sJobInspectionOver )
      Coil( #qJobInspectionOver )
   END_RUNG
   // the same network as SCL:
   #qVisionOnline := true AND #iqInsight_Camera.Vision_Input.iOnline;
   #qVisionOfflineReason1 := true AND #iqInsight_Camera.Vision_Input."iOffline Reason_0";
   #qVisionOfflineReason2 := true AND #iqInsight_Camera.Vision_Input."iOffline Reason_1";
   #qVisionOfflineReason3 := true AND #iqInsight_Camera.Vision_Input."iOffline Reason_2";
   #sJobInspectionOver := true AND #iStartInspection AND (#sJobPass OR #sJobFail);
   #qJobInspectionOver := true AND #sJobInspectionOver;
END_REGION

REGION Network 33: Errors
   // Errors: 
   // qErrTriggerTimeOut: Tigger TimeOut Error Occured
   // qErrAcquiringTimeout: Acquiring TimeOut Error Occured
   // qErrTriggerEnableTimeout: Trigger Enable TimeOut Occured
   // Errors: 
   // qErrTriggerTimeOut: Trigger TimeOut Error Occured
   // qErrAcquiringTimeout: Acquiring TimeOut Error Occured
   // qErrTriggerEnableTimeout: Trigger Enable TimeOut Occured
   // qErrJobSelection: Job selection Error
   // qBothStartOn: Both Start are ON
   RUNG wire#powerrail
      Contact( true )
      Contact( #iAutorunning )
      wire#w1
      Contact( #iStartInspection )
      wire#w2
      Contact( #TriggerTimeout.Q )
      wire#w3
      Coil( #sErrTriggerTimeOut )
   END_RUNG
   RUNG wire#w2
      Contact( #sErrTriggerTimeOut )
      I_Contact( #iResetFault )
   END_RUNG wire#w3
   RUNG wire#w2
      Contact( #AcquiringTimeOut.Q )
      wire#w4
      Coil( #sErrAcquiringTimeOut )
   END_RUNG
   RUNG wire#w2
      Contact( #sErrAcquiringTimeOut )
      I_Contact( #iResetFault )
   END_RUNG wire#w4
   RUNG wire#w2
      Contact( #TriggerEnableTimeout.Q )
      wire#w5
      Coil( #sErrTriggerEnableTimeout )
   END_RUNG
   RUNG wire#w2
      Contact( #sErrTriggerEnableTimeout )
      I_Contact( #iResetFault )
   END_RUNG wire#w5
   RUNG wire#w1
      Contact( #sProgramEcho.Q )
      { S7_Templates := "SrcType := Int" } NE_Contact(in1 := #iJobID, in2 := #sVisionInputCmdControlIP)
      I_Contact( #sJobSelectionOver )
      wire#w6
      Coil( #sErrJobSelection )
   END_RUNG
   RUNG wire#w1
      Contact( #sErrJobSelection )
      I_Contact( #iResetFault )
   END_RUNG wire#w6
   RUNG wire#w1
      Contact( #iStartInspection )
      Contact( #iStartJobSelection )
      wire#w7
      Coil( #sBothStartOn )
   END_RUNG
   RUNG wire#w1
      Contact( #sBothStartOn )
      I_Contact( #iResetFault )
   END_RUNG wire#w7
   // the same network as SCL:
   #_w1 := true AND #iAutorunning;
   #_w2 := #_w1 AND #iStartInspection;
   #sErrTriggerTimeOut := #_w2 AND (#TriggerTimeout.Q OR (#sErrTriggerTimeOut AND NOT #iResetFault));
   #sErrAcquiringTimeOut := #_w2 AND (#AcquiringTimeOut.Q OR (#sErrAcquiringTimeOut AND NOT #iResetFault));
   #sErrTriggerEnableTimeout := #_w2 AND (#TriggerEnableTimeout.Q OR (#sErrTriggerEnableTimeout AND NOT #iResetFault));
   #sErrJobSelection := #_w1 AND ((#sProgramEcho.Q AND (#iJobID <> #sVisionInputCmdControlIP) AND NOT #sJobSelectionOver) OR (#sErrJobSelection AND NOT #iResetFault));
   #sBothStartOn := #_w1 AND ((#iStartInspection AND #iStartJobSelection) OR (#sBothStartOn AND NOT #iResetFault));
END_REGION

REGION Network 34: Stat bit Error Mapping / Output mapping using Stat Bit
   // Stat bit Error Mapping / Output mapping using Stat Bit
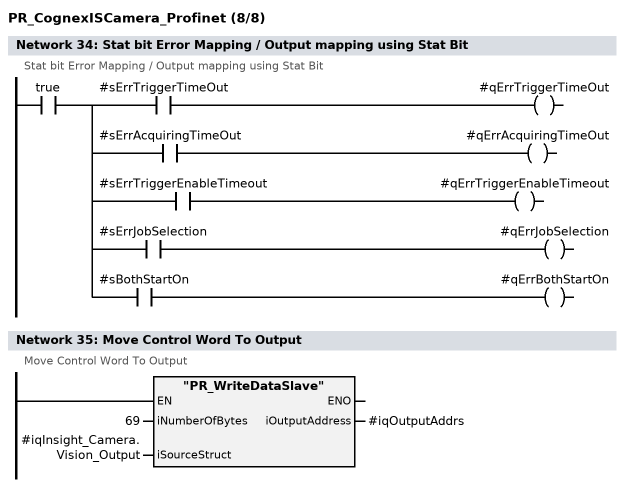
   RUNG wire#powerrail
      Contact( true )
      wire#w1
      Contact( #sErrTriggerTimeOut )
      Coil( #qErrTriggerTimeOut )
   END_RUNG
   RUNG wire#w1
      Contact( #sErrAcquiringTimeOut )
      Coil( #qErrAcquiringTimeOut )
   END_RUNG
   RUNG wire#w1
      Contact( #sErrTriggerEnableTimeout )
      Coil( #qErrTriggerEnableTimeout )
   END_RUNG
   RUNG wire#w1
      Contact( #sErrJobSelection )
      Coil( #qErrJobSelection )
   END_RUNG
   RUNG wire#w1
      Contact( #sBothStartOn )
      Coil( #qErrBothStartOn )
   END_RUNG
   // the same network as SCL:
   #qErrTriggerTimeOut := true AND #sErrTriggerTimeOut;
   #qErrAcquiringTimeOut := true AND #sErrAcquiringTimeOut;
   #qErrTriggerEnableTimeout := true AND #sErrTriggerEnableTimeout;
   #qErrJobSelection := true AND #sErrJobSelection;
   #qErrBothStartOn := true AND #sBothStartOn;
END_REGION

REGION Network 35: Move Control Word To Output
   // Move Control Word To Output
   RUNG wire#powerrail
      "PR_WriteDataSlave"(iNumberOfBytes := 69, iSourceStruct := #iqInsight_Camera.Vision_Output, iOutputAddress => #iqOutputAddrs)
   END_RUNG
   // the same network as SCL:
   "PR_WriteDataSlave"(iNumberOfBytes := 69,
                       iSourceStruct := #iqInsight_Camera.Vision_Output,
                       iOutputAddress => #iqOutputAddrs);
END_REGION
END_FUNCTION_BLOCK

FUNCTION_BLOCK "PR_CognexIS28xx_Profi"   // FB496, LAD
TITLE = PR_CognexIS28xx_Profi
{ S7_Optimized_Access := 'TRUE' }
AUTHOR : MS
FAMILY : WiproPari
NAME : S21006022015
VERSION : 0.3
   VAR_INPUT
      iInsightCamera_Input : "UDT_IS28xx_To_Plc";   // Connect Camera Input
      iResetFault : Bool;   // Reset Fault Input
      iModuleReset : Bool;   // Connect Module reset Signal to this pin
      iAutorunning : Bool;   // Autorunning Input
      iStartJobSelection : Bool;   // start job selection
      iStartInspection : Bool;   // start inspection
      iJobID : Int;   // job id
      iUserData : Array[1..60] of Byte;   // Enter user data which is send to cognex camera/controller
      iTriggerEnableTimeoutTime : Time;   // Trigger Enable TimeOut Time Delay
      iTriggerTimeoutTime : Time;   // Trigger TimeOut Time Delay
      iAcquiringTimeOutTime : Time;   // Acquiring TimeOut Time Delay
      iPrgmNoTimeOut : Time;   // Timeout for program echo received from camera
      iFeedbackTimeOut : Time;   // Feedback time out time
   END_VAR
   VAR_OUTPUT
      qInsightCamera_Output : "UDT_Plc_To_IS28xx";   // Connect Camera Output
      qJobPass : Bool;   // Job Pass In Inspection
      qJobFail : Bool;   // Job Failed In Inspection
      qJobSelectionOver : Bool;   // job selection over
      qJobInspectionOver : Bool;   // Inspection Over Output
      qVisionOnline : Bool;   // Insight Vision Is In Online
      qVisionOfflineReason1 : Bool;   // Insight Vision Offline Due To: The vision system's job is being modified
      qVisionOfflineReason2 : Bool;   // Insight Vision Offline Due To: A discrete signal is holding the vision system Offline
      qVisionOfflineReason3 : Bool;   // Insight Vision Offline Due To: A communications protocol is holding the vision system Offline
      qErrBothStartOn : Bool;   // both start on
      qErrJobSelection : Bool;   // error job selection
      qErrTriggerEnableTimeout : Bool;   // Trigger Enable TimeOut Error
      qErrTriggerTimeOut : Bool;   // Trigger TimeOut Error
      qErrAcquiringTimeOut : Bool;   // Acquiring TimeOut Error
      qErrJobIDEchoMismatch : Bool;   // Job Id Echo mismatch Error
      qErrSetUserDataAckNtRcvd : Bool;   // Set user data ack not received within time
      qMsgJobIDMismatch : Bool;   // Selected Job ID & Running JOB ID not matched message
      qInspectionResult : Array[1..60] of Byte;   // Inspection Result Data
   END_VAR
   VAR_IN_OUT
      iqRunningJobID : Int;   // It Shows running Job ID
   END_VAR
   VAR
      sResetFaults : Bool;
      sInspectionComplete : Bool;
      sJobPass : Bool;
      sJobFail : Bool;
      sJobLoadcompleted : Bool;
      sJobSelectionOver : Bool;
      sJobInspectionOver : Bool;
      sVisionOutput_Trigger : Bool;
      sInitialPulse : Bool;
      sExposureTimerStar1 : Bool;
      sExposureTimerStart : Bool;
      sPulse : Array[0..7] of Bool;
      sVisionInputCmdControlIP : Int;
      sTriggerEnableTimeoutTime : Time;
      sTriggerTimeoutTime : Time;
      sAcquiringTimeOutTime : Time;
      TriggerTimeout : TON_TIME;
      TriggerEnableTimeout : TON_TIME;
      AcquiringTimeOut : TON_TIME;
      ResultTimer : TON_TIME;
      sExposureTimer : TON_TIME;
      sTriggerResetTimer : TON_TIME;
      sPrgmNoTimeOut : Time;
      sPrgmNumTimer : TON_TIME;
      sSetUserDataAckTimer : TON_TIME;
      sFeedbackTimeOut : Time;
   END_VAR
   VAR_TEMP   // added for the SCL form of the ladder/FBD networks
      _w1 : Bool;
      _w2 : Bool;
      _w3 : Bool;
      _w4 : Bool;
      _w5 : Bool;
   END_VAR
BEGIN

REGION Network 1: Header
   // ==============================================================================
   //  Company: Precision Automation & Robotics India Ltd. 
   // ------------------------------------------------------------------------------
   //  Item Code: S21006022015
   //  Author/Created by: Manoj Sonawane
   //  Reviewed/Checked by: Sandip.c
   //  First Release on: 19-07-24
   //  Latest update on:11-03-25
   // ------------------------------------------------------------------------------
   //  Tested with: CPU firmware, model or simulator testing
   //  Engineering/Editor: TIA Portal V17
   // ------------------------------------------------------------------------------
   //  Restrictions:
   //  Dependencies/Requirements:
   //  1. "UDT_IS28xx_To_Plc"
   //  2. "UDT_Plc_To_IS28xx"
   // ------------------------------------------------------------------------------
   //  Change Log:
   //  Ver.	Date		Changed by		Details of changes
   //  1.0	 19-07-24                 Manoj Sonawane            	First release version
   // 1.1              30-09-24                 Harshal Gharmode                         Modify as per shop floor testing
   // 1.2              11-03-25                 Swapnil Asule                                  Remove retry count logic & update                                                                                                                         data Inspection logic
   // ------------------------------------------------------------------------------
   //  Functionality:  : The Cognex In-Sight® 2801 vision system communicates with the Siemence s7-15xx series PLC over Profinet protocol.The main functionality of this block is provided for the user can change the job ID according to their needs and get the inspection result data of Job ID.
   // 
   // 
   //  Inputs
   // iInsightCamera_Input	"UDT_IS28xx_To_Plc"
   // iResetFault	Bool
   // iModuleReset	Bool
   // iAutorunning	Bool
   // iStartJobSelection	Bool
   // iStartInspection	Bool
   // iJobID	Int
   // iUserData	Array[1..60] of Byte
   // iTriggerEnableTimeoutTime	Time
   // iTriggerTimeoutTime	Time
   // iAcquiringTimeOutTime	Time
   // iPrgmNoTimeOut	Time
   // iFeedbackTimeOut	Time
   // 
   //  Outputs
   //  qInsightCamera_Output	"UDT_Plc_To_IS28xx"
   // qJobPass	Bool
   // qJobFail	Bool
   // qJobSelectionOver	Bool
   // qJobInspectionOver	Bool
   // qVisionOnline	Bool
   // qVisionOfflineReason1	Bool
   // qVisionOfflineReason2	Bool
   // qVisionOfflineReason3	Bool
   // qErrBothStartOn	Bool
   // qErrJobSelection	Bool
   // qErrTriggerEnableTimeout	Bool
   // qErrTriggerTimeOut	Bool
   // qErrAcquiringTimeOut	Bool
   // qErrJobIDEchoMismatch	Bool
   // qErrSetUserDataAckNtRcvd	Bool
   // qMsgJobIDMismatch	Bool
   // qInspectionResult	Array[1..60] of Byte
   // 
   //  In-outs
   //  iqRunningJobID	Int
   // ------------------------------------------------------------------------------
   //  Errors reported:
   //  1.qErrTriggerTimeO : Error trigger timeout
   //  2. qErrAcquiringTimeOut;Acquiring Time Out
   //  3. qErrTriggerEnableTimeout:Trigger Enable Time Out
   //  4. qErrJobSelection: Job selection error
   //  5. qErrBothStartOn: Start Inspection & Start Job Selection command are active at same time
   //  6. qErrJobIDEchoMismatch: Set Job ID & its echo is not matched
   //  7. qErrSetUserDataAckNtRcvd: Set user data acknowldge not recived within the defined time.
   // 
   //  Messages reported:
   //   1. qMsgJobIDMismatch: Set Job ID & running JOB ID is not matched
   // ==============================================================================
END_REGION

REGION Network 2: Reset Faults
   // Reset Faults
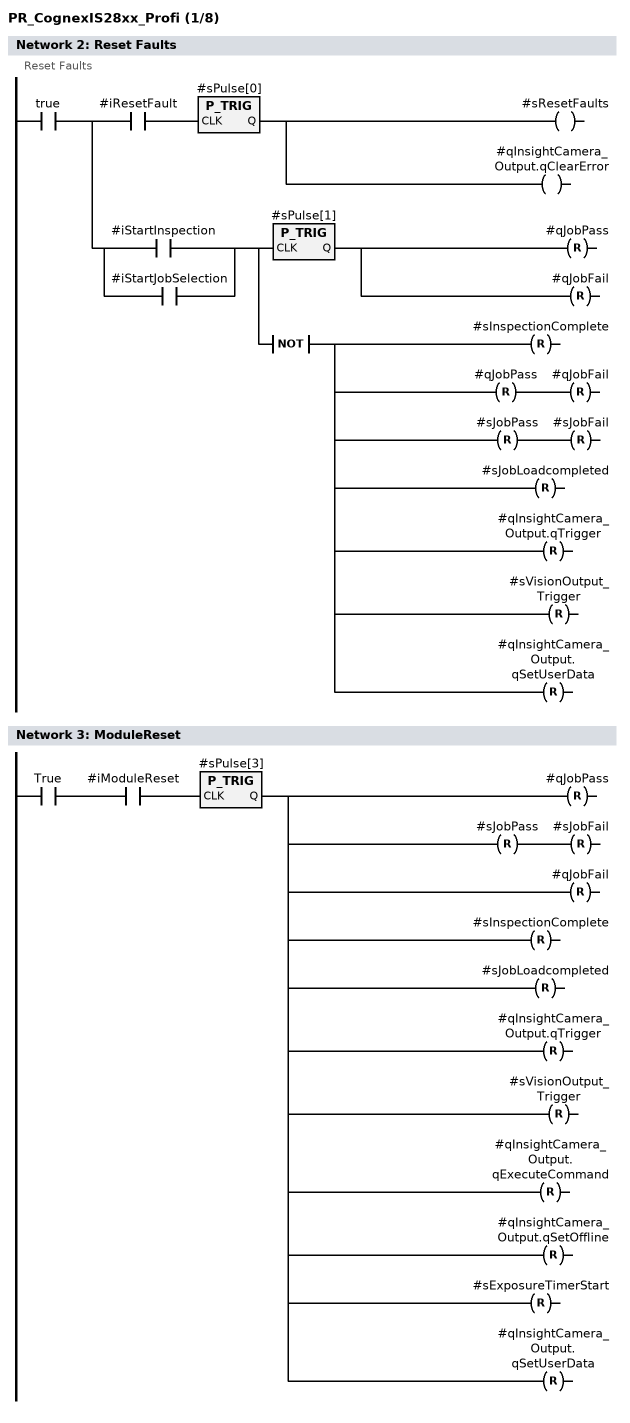
   RUNG wire#powerrail
      Contact( true )
      wire#w1
      Contact( #iResetFault )
      P_Trig( #sPulse[0] )
      wire#w2
      Coil( #sResetFaults )
   END_RUNG
   RUNG wire#w2
      Coil( #qInsightCamera_Output.qClearError )
   END_RUNG
   RUNG wire#w1
      Contact( #iStartInspection )
      wire#w3
      P_Trig( #sPulse[1] )
      wire#w4
      R_Coil( #qJobPass )
   END_RUNG
   RUNG wire#w1
      Contact( #iStartJobSelection )
   END_RUNG wire#w3
   RUNG wire#w4
      R_Coil( #qJobFail )
   END_RUNG
   RUNG wire#w3
      Not()
      wire#w5
      R_Coil( #sInspectionComplete )
   END_RUNG
   RUNG wire#w5
      R_Coil( #qJobPass )
      R_Coil( #qJobFail )
   END_RUNG
   RUNG wire#w5
      R_Coil( #sJobPass )
      R_Coil( #sJobFail )
   END_RUNG
   RUNG wire#w5
      R_Coil( #sJobLoadcompleted )
   END_RUNG
   RUNG wire#w5
      R_Coil( #qInsightCamera_Output.qTrigger )
   END_RUNG
   RUNG wire#w5
      R_Coil( #sVisionOutput_Trigger )
   END_RUNG
   RUNG wire#w5
      R_Coil( #qInsightCamera_Output.qSetUserData )
   END_RUNG
   // the same network as SCL:
   #_w1 := true AND #iResetFault;
   #_w2 := #_w1 AND NOT #sPulse[0];   // rising edge
   #sPulse[0] := #_w1;
   #sResetFaults := #_w2;
   #qInsightCamera_Output.qClearError := #_w2;
   #_w3 := true AND (#iStartInspection OR #iStartJobSelection);
   #_w4 := #_w3 AND NOT #sPulse[1];   // rising edge
   #sPulse[1] := #_w3;
   IF #_w4 THEN
       #qJobPass := FALSE;
       #qJobFail := FALSE;
   END_IF;
   IF NOT #_w3 THEN
       #sInspectionComplete := FALSE;
       #qJobPass := FALSE;
       #qJobFail := FALSE;
       #sJobPass := FALSE;
       #sJobFail := FALSE;
       #sJobLoadcompleted := FALSE;
       #qInsightCamera_Output.qTrigger := FALSE;
       #sVisionOutput_Trigger := FALSE;
       #qInsightCamera_Output.qSetUserData := FALSE;
   END_IF;
END_REGION

REGION Network 3: ModuleReset
   RUNG wire#powerrail
      Contact( True )
      Contact( #iModuleReset )
      P_Trig( #sPulse[3] )
      wire#w1
      R_Coil( #qJobPass )
   END_RUNG
   RUNG wire#w1
      R_Coil( #sJobPass )
      R_Coil( #sJobFail )
   END_RUNG
   RUNG wire#w1
      R_Coil( #qJobFail )
   END_RUNG
   RUNG wire#w1
      R_Coil( #sInspectionComplete )
   END_RUNG
   RUNG wire#w1
      R_Coil( #sJobLoadcompleted )
   END_RUNG
   RUNG wire#w1
      R_Coil( #qInsightCamera_Output.qTrigger )
   END_RUNG
   RUNG wire#w1
      R_Coil( #sVisionOutput_Trigger )
   END_RUNG
   RUNG wire#w1
      R_Coil( #qInsightCamera_Output.qExecuteCommand )
   END_RUNG
   RUNG wire#w1
      R_Coil( #qInsightCamera_Output.qSetOffline )
   END_RUNG
   RUNG wire#w1
      R_Coil( #sExposureTimerStart )
   END_RUNG
   RUNG wire#w1
      R_Coil( #qInsightCamera_Output.qSetUserData )
   END_RUNG
   // the same network as SCL:
   #_w1 := True AND #iModuleReset;
   #_w2 := #_w1 AND NOT #sPulse[3];   // rising edge
   #sPulse[3] := #_w1;
   IF #_w2 THEN
       #qJobPass := FALSE;
       #sJobPass := FALSE;
       #sJobFail := FALSE;
       #qJobFail := FALSE;
       #sInspectionComplete := FALSE;
       #sJobLoadcompleted := FALSE;
       #qInsightCamera_Output.qTrigger := FALSE;
       #sVisionOutput_Trigger := FALSE;
       #qInsightCamera_Output.qExecuteCommand := FALSE;
       #qInsightCamera_Output.qSetOffline := FALSE;
       #sExposureTimerStart := FALSE;
       #qInsightCamera_Output.qSetUserData := FALSE;
   END_IF;
END_REGION

REGION Network 4: Time out validation
   // Time out validation 1. Trigger enable time out
   // 2. Trigger time out
   // 3. Acquiring TimeOut Time
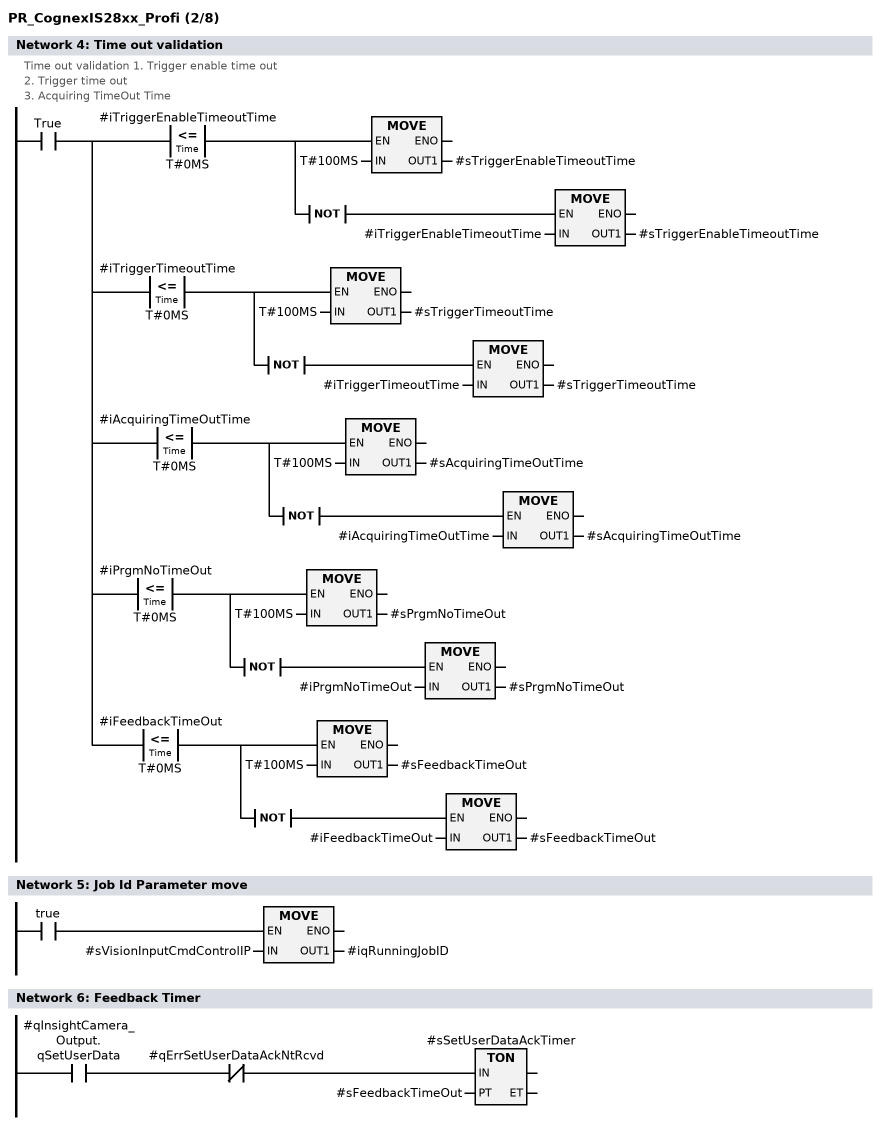
   RUNG wire#powerrail
      Contact( True )
      wire#w1
      { S7_Templates := "SrcType := Time" } LE_Contact(in1 := #iTriggerEnableTimeoutTime, in2 := T#0MS)
      wire#w2
      Move(in := T#100MS, out1 => #sTriggerEnableTimeoutTime)
   END_RUNG
   RUNG wire#w2
      Not()
      Move(in := #iTriggerEnableTimeoutTime, out1 => #sTriggerEnableTimeoutTime)
   END_RUNG
   RUNG wire#w1
      { S7_Templates := "SrcType := Time" } LE_Contact(in1 := #iTriggerTimeoutTime, in2 := T#0MS)
      wire#w3
      Move(in := T#100MS, out1 => #sTriggerTimeoutTime)
   END_RUNG
   RUNG wire#w3
      Not()
      Move(in := #iTriggerTimeoutTime, out1 => #sTriggerTimeoutTime)
   END_RUNG
   RUNG wire#w1
      { S7_Templates := "SrcType := Time" } LE_Contact(in1 := #iAcquiringTimeOutTime, in2 := T#0MS)
      wire#w4
      Move(in := T#100MS, out1 => #sAcquiringTimeOutTime)
   END_RUNG
   RUNG wire#w4
      Not()
      Move(in := #iAcquiringTimeOutTime, out1 => #sAcquiringTimeOutTime)
   END_RUNG
   RUNG wire#w1
      { S7_Templates := "SrcType := Time" } LE_Contact(in1 := #iPrgmNoTimeOut, in2 := T#0MS)
      wire#w5
      Move(in := T#100MS, out1 => #sPrgmNoTimeOut)
   END_RUNG
   RUNG wire#w5
      Not()
      Move(in := #iPrgmNoTimeOut, out1 => #sPrgmNoTimeOut)
   END_RUNG
   RUNG wire#w1
      { S7_Templates := "SrcType := Time" } LE_Contact(in1 := #iFeedbackTimeOut, in2 := T#0MS)
      wire#w6
      Move(in := T#100MS, out1 => #sFeedbackTimeOut)
   END_RUNG
   RUNG wire#w6
      Not()
      Move(in := #iFeedbackTimeOut, out1 => #sFeedbackTimeOut)
   END_RUNG
   // the same network as SCL:
   #_w1 := True AND (#iTriggerEnableTimeoutTime <= T#0MS);
   IF #_w1 THEN #sTriggerEnableTimeoutTime := T#100MS; END_IF;
   IF NOT #_w1 THEN #sTriggerEnableTimeoutTime := #iTriggerEnableTimeoutTime; END_IF;
   #_w2 := True AND (#iTriggerTimeoutTime <= T#0MS);
   IF #_w2 THEN #sTriggerTimeoutTime := T#100MS; END_IF;
   IF NOT #_w2 THEN #sTriggerTimeoutTime := #iTriggerTimeoutTime; END_IF;
   #_w3 := True AND (#iAcquiringTimeOutTime <= T#0MS);
   IF #_w3 THEN #sAcquiringTimeOutTime := T#100MS; END_IF;
   IF NOT #_w3 THEN #sAcquiringTimeOutTime := #iAcquiringTimeOutTime; END_IF;
   #_w4 := True AND (#iPrgmNoTimeOut <= T#0MS);
   IF #_w4 THEN #sPrgmNoTimeOut := T#100MS; END_IF;
   IF NOT #_w4 THEN #sPrgmNoTimeOut := #iPrgmNoTimeOut; END_IF;
   #_w5 := True AND (#iFeedbackTimeOut <= T#0MS);
   IF #_w5 THEN #sFeedbackTimeOut := T#100MS; END_IF;
   IF NOT #_w5 THEN #sFeedbackTimeOut := #iFeedbackTimeOut; END_IF;
END_REGION

REGION Network 5: Job Id Parameter move
   RUNG wire#powerrail
      Contact( true )
      Move(in := #sVisionInputCmdControlIP, out1 => #iqRunningJobID)
   END_RUNG
   // the same network as SCL:
   IF true THEN #iqRunningJobID := #sVisionInputCmdControlIP; END_IF;
END_REGION

REGION Network 6: Feedback Timer
   #sSetUserDataAckTimer(IN := #qInsightCamera_Output.qSetUserData AND NOT #qErrSetUserDataAckNtRcvd,   // TON
                         PT := #sFeedbackTimeOut);
END_REGION

REGION Network 7: UserData
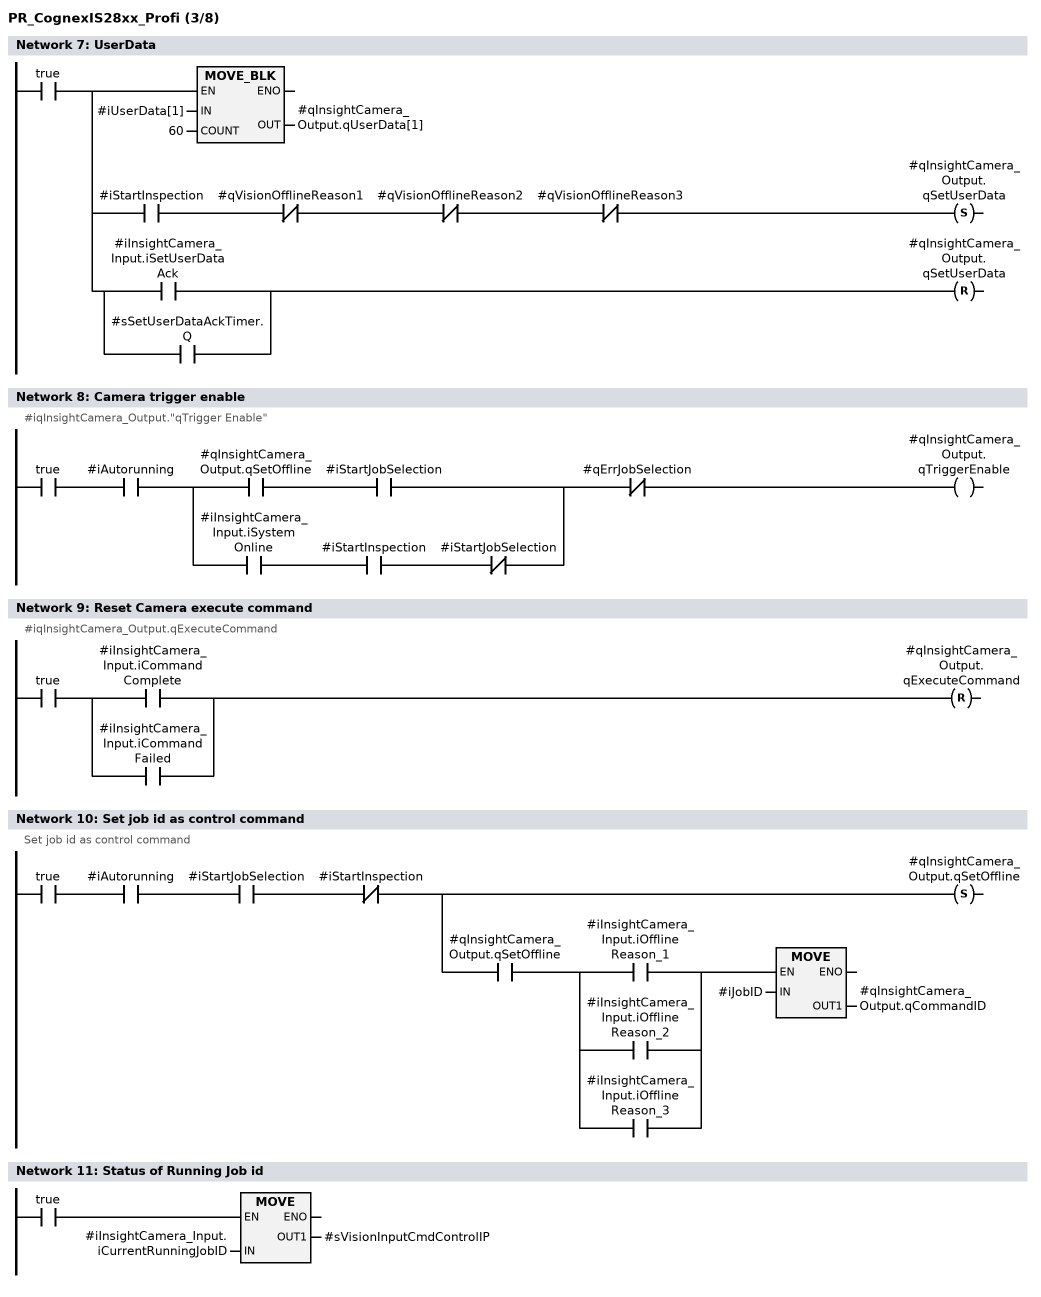
   IF true THEN
       MOVE_BLK(IN := #iUserData[1], COUNT := 60, OUT => #qInsightCamera_Output.qUserData[1]);
   END_IF;
   IF true AND #iStartInspection AND NOT #qVisionOfflineReason1 AND NOT #qVisionOfflineReason2 AND NOT #qVisionOfflineReason3 THEN
       #qInsightCamera_Output.qSetUserData := TRUE;
   END_IF;
   IF true AND (#iInsightCamera_Input.iSetUserDataAck OR #sSetUserDataAckTimer.Q) THEN
       #qInsightCamera_Output.qSetUserData := FALSE;
   END_IF;
END_REGION

REGION Network 8: Camera trigger enable
   // #iqInsightCamera_Output."qTrigger Enable"
   RUNG wire#powerrail
      Contact( true )
      Contact( #iAutorunning )
      wire#w1
      Contact( #qInsightCamera_Output.qSetOffline )
      Contact( #iStartJobSelection )
      wire#w2
      I_Contact( #qErrJobSelection )
      Coil( #qInsightCamera_Output.qTriggerEnable )
   END_RUNG
   RUNG wire#w1
      Contact( #iInsightCamera_Input.iSystemOnline )
      Contact( #iStartInspection )
      I_Contact( #iStartJobSelection )
   END_RUNG wire#w2
   // the same network as SCL:
   #qInsightCamera_Output.qTriggerEnable := true AND #iAutorunning AND ((#qInsightCamera_Output.qSetOffline AND #iStartJobSelection) OR (#iInsightCamera_Input.iSystemOnline AND #iStartInspection AND NOT #iStartJobSelection)) AND NOT #qErrJobSelection;
END_REGION

REGION Network 9: Reset Camera execute command
   // #iqInsightCamera_Output.qExecuteCommand
   RUNG wire#powerrail
      Contact( true )
      wire#w1
      Contact( #iInsightCamera_Input.iCommandComplete )
      wire#w2
      R_Coil( #qInsightCamera_Output.qExecuteCommand )
   END_RUNG
   RUNG wire#w1
      Contact( #iInsightCamera_Input.iCommandFailed )
   END_RUNG wire#w2
   // the same network as SCL:
   IF true AND (#iInsightCamera_Input.iCommandComplete OR #iInsightCamera_Input.iCommandFailed) THEN
       #qInsightCamera_Output.qExecuteCommand := FALSE;
   END_IF;
END_REGION

REGION Network 10: Set job id as control command
   // Set job id as control command
   RUNG wire#powerrail
      Contact( true )
      Contact( #iAutorunning )
      Contact( #iStartJobSelection )
      I_Contact( #iStartInspection )
      wire#w1
      S_Coil( #qInsightCamera_Output.qSetOffline )
   END_RUNG
   RUNG wire#w1
      Contact( #qInsightCamera_Output.qSetOffline )
      wire#w2
      Contact( #iInsightCamera_Input.iOfflineReason_1 )
      wire#w3
      Move(in := #iJobID, out1 => #qInsightCamera_Output.qCommandID)
   END_RUNG
   RUNG wire#w2
      Contact( #iInsightCamera_Input.iOfflineReason_2 )
   END_RUNG wire#w3
   RUNG wire#w2
      Contact( #iInsightCamera_Input.iOfflineReason_3 )
   END_RUNG wire#w3
   // the same network as SCL:
   #_w1 := true AND #iAutorunning AND #iStartJobSelection AND NOT #iStartInspection;
   IF #_w1 THEN #qInsightCamera_Output.qSetOffline := TRUE; END_IF;
   IF #_w1 AND #qInsightCamera_Output.qSetOffline AND (#iInsightCamera_Input.iOfflineReason_1 OR #iInsightCamera_Input.iOfflineReason_2 OR #iInsightCamera_Input.iOfflineReason_3) THEN
       #qInsightCamera_Output.qCommandID := #iJobID;
   END_IF;
END_REGION

REGION Network 11: Status of Running Job id
   RUNG wire#powerrail
      Contact( true )
      Move(in := #iInsightCamera_Input.iCurrentRunningJobID, out1 => #sVisionInputCmdControlIP)
   END_RUNG
   // the same network as SCL:
   IF true THEN #sVisionInputCmdControlIP := #iInsightCamera_Input.iCurrentRunningJobID; END_IF;
END_REGION

REGION Network 12: Set Execute command as per Job selection
   // Set Execute command as per Job selection
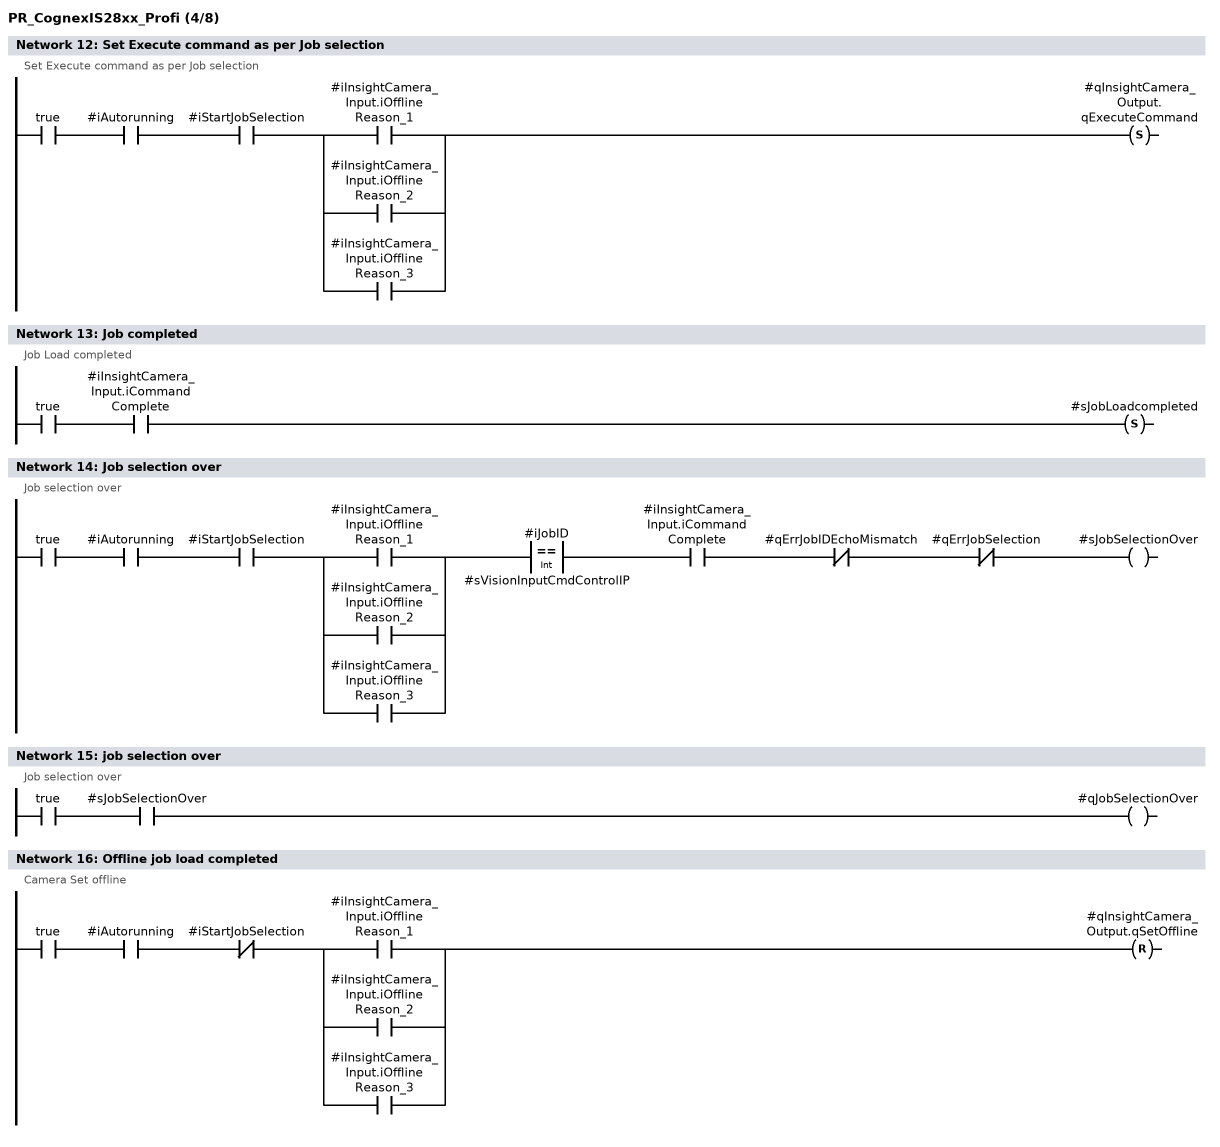
   RUNG wire#powerrail
      Contact( true )
      Contact( #iAutorunning )
      Contact( #iStartJobSelection )
      wire#w1
      Contact( #iInsightCamera_Input.iOfflineReason_1 )
      wire#w2
      S_Coil( #qInsightCamera_Output.qExecuteCommand )
   END_RUNG
   RUNG wire#w1
      Contact( #iInsightCamera_Input.iOfflineReason_2 )
   END_RUNG wire#w2
   RUNG wire#w1
      Contact( #iInsightCamera_Input.iOfflineReason_3 )
   END_RUNG wire#w2
   // the same network as SCL:
   IF true AND #iAutorunning AND #iStartJobSelection AND (#iInsightCamera_Input.iOfflineReason_1 OR #iInsightCamera_Input.iOfflineReason_2 OR #iInsightCamera_Input.iOfflineReason_3) THEN
       #qInsightCamera_Output.qExecuteCommand := TRUE;
   END_IF;
END_REGION

REGION Network 13: Job completed
   // Job Load completed
   RUNG wire#powerrail
      Contact( true )
      Contact( #iInsightCamera_Input.iCommandComplete )
      S_Coil( #sJobLoadcompleted )
   END_RUNG
   // the same network as SCL:
   IF true AND #iInsightCamera_Input.iCommandComplete THEN #sJobLoadcompleted := TRUE; END_IF;
END_REGION

REGION Network 14: Job selection over
   // Job selection over
   RUNG wire#powerrail
      Contact( true )
      Contact( #iAutorunning )
      Contact( #iStartJobSelection )
      wire#w1
      Contact( #iInsightCamera_Input.iOfflineReason_1 )
      wire#w2
      { S7_Templates := "SrcType := Int" } EQ_Contact(in1 := #iJobID, in2 := #sVisionInputCmdControlIP)
      Contact( #iInsightCamera_Input.iCommandComplete )
      I_Contact( #qErrJobIDEchoMismatch )
      I_Contact( #qErrJobSelection )
      Coil( #sJobSelectionOver )
   END_RUNG
   RUNG wire#w1
      Contact( #iInsightCamera_Input.iOfflineReason_2 )
   END_RUNG wire#w2
   RUNG wire#w1
      Contact( #iInsightCamera_Input.iOfflineReason_3 )
   END_RUNG wire#w2
   // the same network as SCL:
   #sJobSelectionOver := true AND #iAutorunning AND #iStartJobSelection AND (#iInsightCamera_Input.iOfflineReason_1 OR #iInsightCamera_Input.iOfflineReason_2 OR #iInsightCamera_Input.iOfflineReason_3) AND (#iJobID = #sVisionInputCmdControlIP) AND #iInsightCamera_Input.iCommandComplete AND NOT #qErrJobIDEchoMismatch AND NOT #qErrJobSelection;
END_REGION

REGION Network 15: job selection over
   // Job selection over
   RUNG wire#powerrail
      Contact( true )
      Contact( #sJobSelectionOver )
      Coil( #qJobSelectionOver )
   END_RUNG
   // the same network as SCL:
   #qJobSelectionOver := true AND #sJobSelectionOver;
END_REGION

REGION Network 16: Offline job load completed
   // Camera Set offline
   RUNG wire#powerrail
      Contact( true )
      Contact( #iAutorunning )
      I_Contact( #iStartJobSelection )
      wire#w1
      Contact( #iInsightCamera_Input.iOfflineReason_1 )
      wire#w2
      R_Coil( #qInsightCamera_Output.qSetOffline )
   END_RUNG
   RUNG wire#w1
      Contact( #iInsightCamera_Input.iOfflineReason_2 )
   END_RUNG wire#w2
   RUNG wire#w1
      Contact( #iInsightCamera_Input.iOfflineReason_3 )
   END_RUNG wire#w2
   // the same network as SCL:
   IF true AND #iAutorunning AND NOT #iStartJobSelection AND (#iInsightCamera_Input.iOfflineReason_1 OR #iInsightCamera_Input.iOfflineReason_2 OR #iInsightCamera_Input.iOfflineReason_3) THEN
       #qInsightCamera_Output.qSetOffline := FALSE;
   END_IF;
END_REGION

REGION Network 17: Trigger Enable
   // Trigger Enable
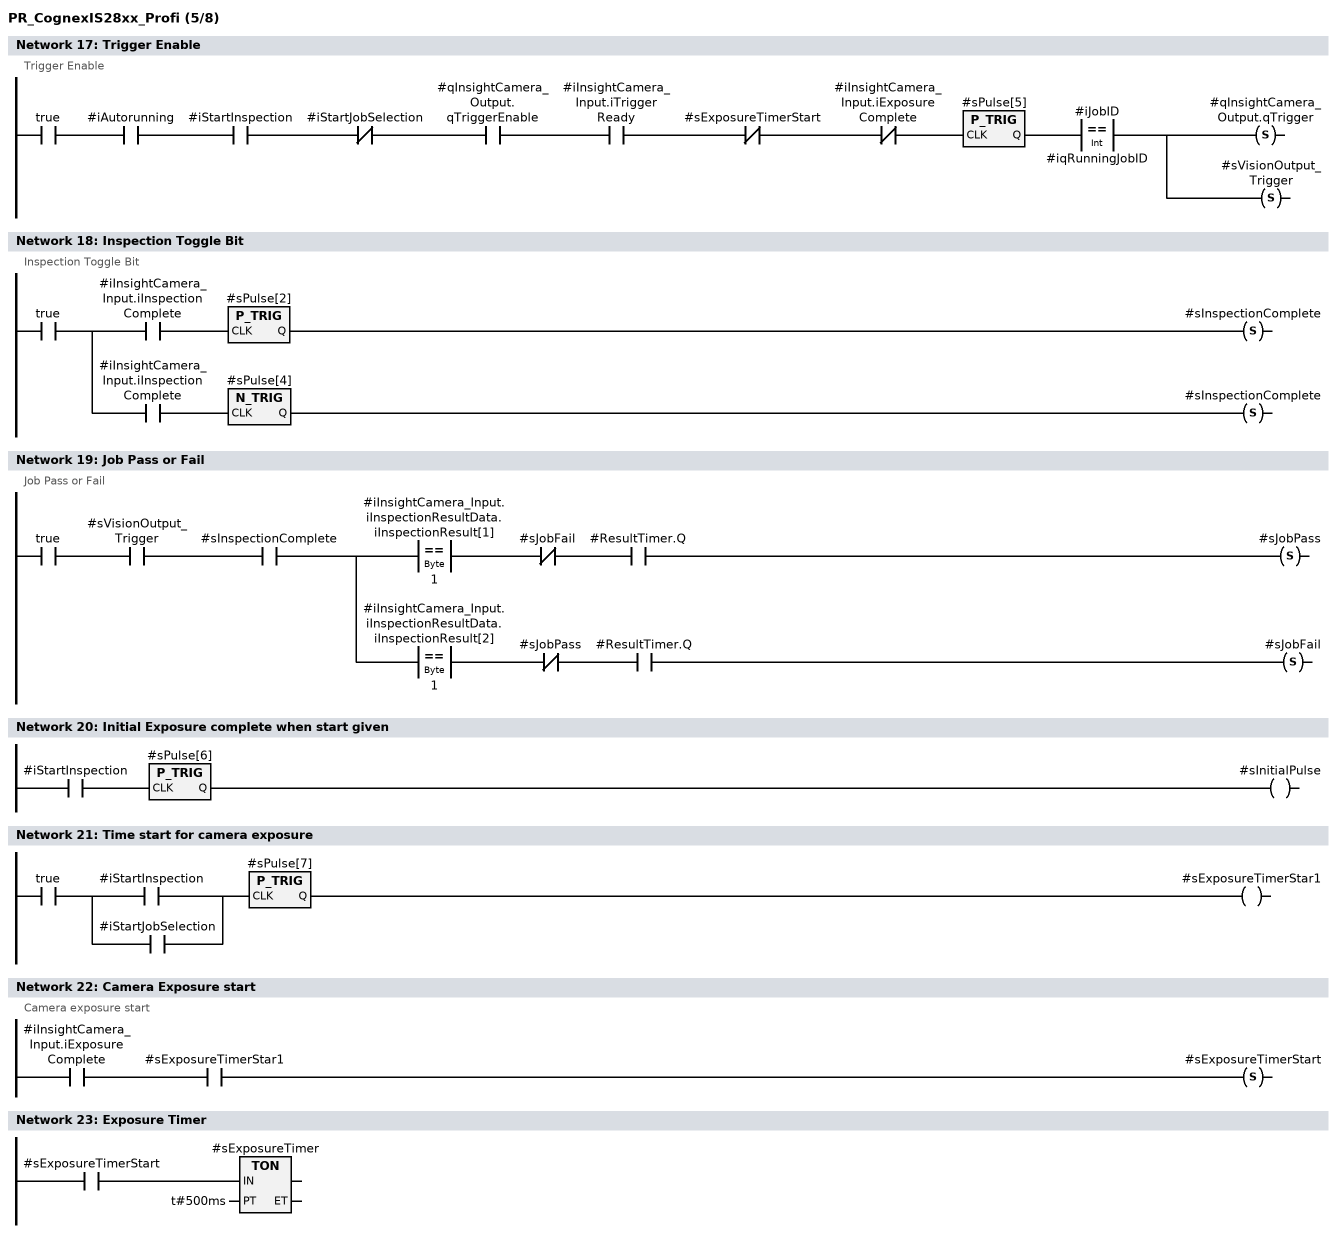
   RUNG wire#powerrail
      Contact( true )
      Contact( #iAutorunning )
      Contact( #iStartInspection )
      I_Contact( #iStartJobSelection )
      Contact( #qInsightCamera_Output.qTriggerEnable )
      Contact( #iInsightCamera_Input.iTriggerReady )
      I_Contact( #sExposureTimerStart )
      I_Contact( #iInsightCamera_Input.iExposureComplete )
      P_Trig( #sPulse[5] )
      { S7_Templates := "SrcType := Int" } EQ_Contact(in1 := #iJobID, in2 := #iqRunningJobID)
      wire#w1
      S_Coil( #qInsightCamera_Output.qTrigger )
   END_RUNG
   RUNG wire#w1
      S_Coil( #sVisionOutput_Trigger )
   END_RUNG
   // the same network as SCL:
   #_w1 := true AND #iAutorunning AND #iStartInspection AND NOT #iStartJobSelection AND #qInsightCamera_Output.qTriggerEnable AND #iInsightCamera_Input.iTriggerReady AND NOT #sExposureTimerStart AND NOT #iInsightCamera_Input.iExposureComplete;
   #_w2 := #_w1 AND NOT #sPulse[5];   // rising edge
   #sPulse[5] := #_w1;
   IF #_w2 AND (#iJobID = #iqRunningJobID) THEN
       #qInsightCamera_Output.qTrigger := TRUE;
       #sVisionOutput_Trigger := TRUE;
   END_IF;
END_REGION

REGION Network 18: Inspection Toggle Bit
   // Inspection Toggle Bit
   RUNG wire#powerrail
      Contact( true )
      wire#w1
      Contact( #iInsightCamera_Input.iInspectionComplete )
      P_Trig( #sPulse[2] )
      S_Coil( #sInspectionComplete )
   END_RUNG
   RUNG wire#w1
      Contact( #iInsightCamera_Input.iInspectionComplete )
      N_Trig( #sPulse[4] )
      S_Coil( #sInspectionComplete )
   END_RUNG
   // the same network as SCL:
   #_w1 := true AND #iInsightCamera_Input.iInspectionComplete;
   #_w2 := #_w1 AND NOT #sPulse[2];   // rising edge
   #sPulse[2] := #_w1;
   IF #_w2 THEN #sInspectionComplete := TRUE; END_IF;
   #_w3 := true AND #iInsightCamera_Input.iInspectionComplete;
   #_w4 := NOT #_w3 AND #sPulse[4];   // falling edge
   #sPulse[4] := #_w3;
   IF #_w4 THEN #sInspectionComplete := TRUE; END_IF;
END_REGION

REGION Network 19: Job Pass or Fail
   // Job Pass or Fail
   RUNG wire#powerrail
      Contact( true )
      Contact( #sVisionOutput_Trigger )
      Contact( #sInspectionComplete )
      wire#w1
      { S7_Templates := "SrcType := Byte" } EQ_Contact(in1 := #iInsightCamera_Input.iInspectionResultData.iInspectionResult[1], in2 := 1)
      I_Contact( #sJobFail )
      Contact( #ResultTimer.Q )
      S_Coil( #sJobPass )
   END_RUNG
   RUNG wire#w1
      { S7_Templates := "SrcType := Byte" } EQ_Contact(in1 := #iInsightCamera_Input.iInspectionResultData.iInspectionResult[2], in2 := 1)
      I_Contact( #sJobPass )
      Contact( #ResultTimer.Q )
      S_Coil( #sJobFail )
   END_RUNG
   // the same network as SCL:
   #_w1 := true AND #sVisionOutput_Trigger AND #sInspectionComplete;
   IF #_w1 AND (#iInsightCamera_Input.iInspectionResultData.iInspectionResult[1] = 1) AND NOT #sJobFail AND #ResultTimer.Q THEN
       #sJobPass := TRUE;
   END_IF;
   IF #_w1 AND (#iInsightCamera_Input.iInspectionResultData.iInspectionResult[2] = 1) AND NOT #sJobPass AND #ResultTimer.Q THEN
       #sJobFail := TRUE;
   END_IF;
END_REGION

REGION Network 20: Initial Exposure complete when start given
   RUNG wire#powerrail
      Contact( #iStartInspection )
      P_Trig( #sPulse[6] )
      Coil( #sInitialPulse )
   END_RUNG
   // the same network as SCL:
   #_w1 := #iStartInspection AND NOT #sPulse[6];   // rising edge
   #sPulse[6] := #iStartInspection;
   #sInitialPulse := #_w1;
END_REGION

REGION Network 21: Time start for camera exposure
   RUNG wire#powerrail
      Contact( true )
      wire#w1
      Contact( #iStartInspection )
      wire#w2
      P_Trig( #sPulse[7] )
      Coil( #sExposureTimerStar1 )
   END_RUNG
   RUNG wire#w1
      Contact( #iStartJobSelection )
   END_RUNG wire#w2
   // the same network as SCL:
   #_w1 := true AND (#iStartInspection OR #iStartJobSelection);
   #_w2 := #_w1 AND NOT #sPulse[7];   // rising edge
   #sPulse[7] := #_w1;
   #sExposureTimerStar1 := #_w2;
END_REGION

REGION Network 22: Camera Exposure start
   // Camera exposure start
   RUNG wire#powerrail
      Contact( #iInsightCamera_Input.iExposureComplete )
      Contact( #sExposureTimerStar1 )
      S_Coil( #sExposureTimerStart )
   END_RUNG
   // the same network as SCL:
   IF #iInsightCamera_Input.iExposureComplete AND #sExposureTimerStar1 THEN
       #sExposureTimerStart := TRUE;
   END_IF;
END_REGION

REGION Network 23: Exposure Timer
   #sExposureTimer(IN := #sExposureTimerStart, PT := t#500ms);   // TON
END_REGION

REGION Network 24: Exposure Timer Complete
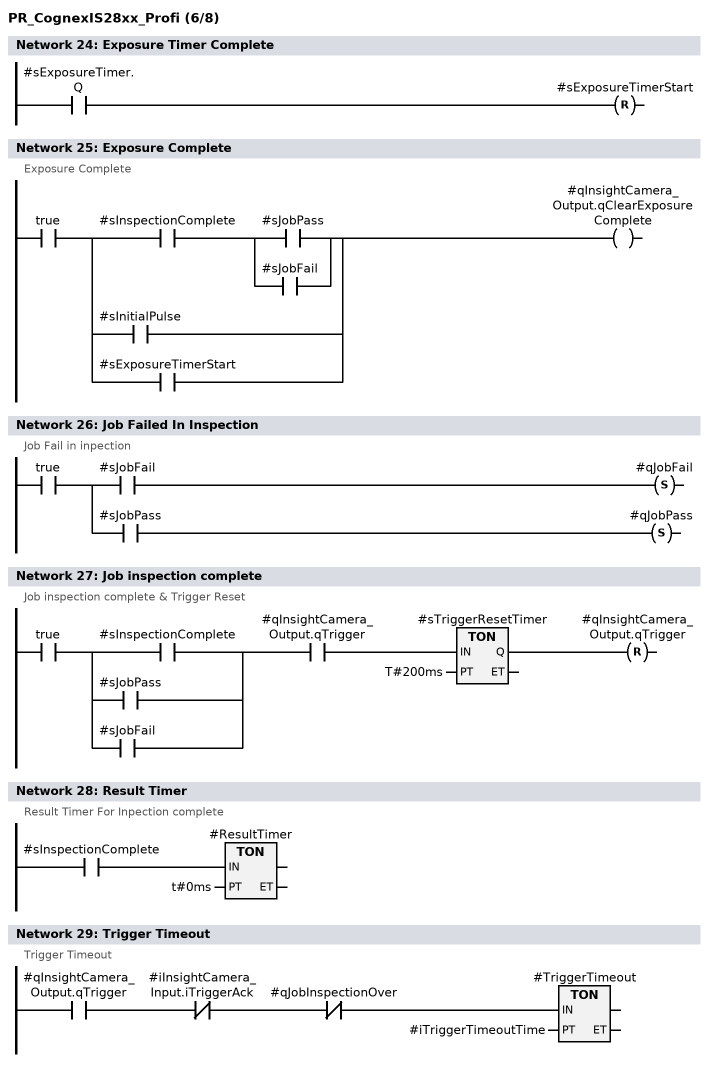
   RUNG wire#powerrail
      Contact( #sExposureTimer.Q )
      R_Coil( #sExposureTimerStart )
   END_RUNG
   // the same network as SCL:
   IF #sExposureTimer.Q THEN #sExposureTimerStart := FALSE; END_IF;
END_REGION

REGION Network 25: Exposure Complete
   // Exposure Complete
   RUNG wire#powerrail
      Contact( true )
      wire#w1
      Contact( #sInspectionComplete )
      wire#w2
      Contact( #sJobPass )
      wire#w3
      Coil( #qInsightCamera_Output.qClearExposureComplete )
   END_RUNG
   RUNG wire#w2
      Contact( #sJobFail )
   END_RUNG wire#w3
   RUNG wire#w1
      Contact( #sInitialPulse )
   END_RUNG wire#w3
   RUNG wire#w1
      Contact( #sExposureTimerStart )
   END_RUNG wire#w3
   // the same network as SCL:
   #qInsightCamera_Output.qClearExposureComplete := true AND ((#sInspectionComplete AND (#sJobPass OR #sJobFail)) OR #sInitialPulse OR #sExposureTimerStart);
END_REGION

REGION Network 26: Job Failed In Inspection
   // Job Fail in inpection
   RUNG wire#powerrail
      Contact( true )
      wire#w1
      Contact( #sJobFail )
      S_Coil( #qJobFail )
   END_RUNG
   RUNG wire#w1
      Contact( #sJobPass )
      S_Coil( #qJobPass )
   END_RUNG
   // the same network as SCL:
   IF true AND #sJobFail THEN #qJobFail := TRUE; END_IF;
   IF true AND #sJobPass THEN #qJobPass := TRUE; END_IF;
END_REGION

REGION Network 27: Job inspection complete
   // Job inspection complete & Trigger Reset
   #sTriggerResetTimer(IN := true AND (#sInspectionComplete OR #sJobPass OR #sJobFail) AND #qInsightCamera_Output.qTrigger,   // TON
                       PT := T#200ms);
   IF #sTriggerResetTimer.Q THEN #qInsightCamera_Output.qTrigger := FALSE; END_IF;
END_REGION

REGION Network 28: Result Timer
   // Result Timer For Inpection complete
   #ResultTimer(IN := #sInspectionComplete, PT := t#0ms);   // TON
END_REGION

REGION Network 29: Trigger Timeout
   // Trigger Timeout
   #TriggerTimeout(IN := #qInsightCamera_Output.qTrigger AND NOT #iInsightCamera_Input.iTriggerAck AND NOT #qJobInspectionOver,   // TON
                   PT := #iTriggerTimeoutTime);
END_REGION

REGION Network 30: Trigger Enable TimeOut
   // Trigger Enable TimeOut
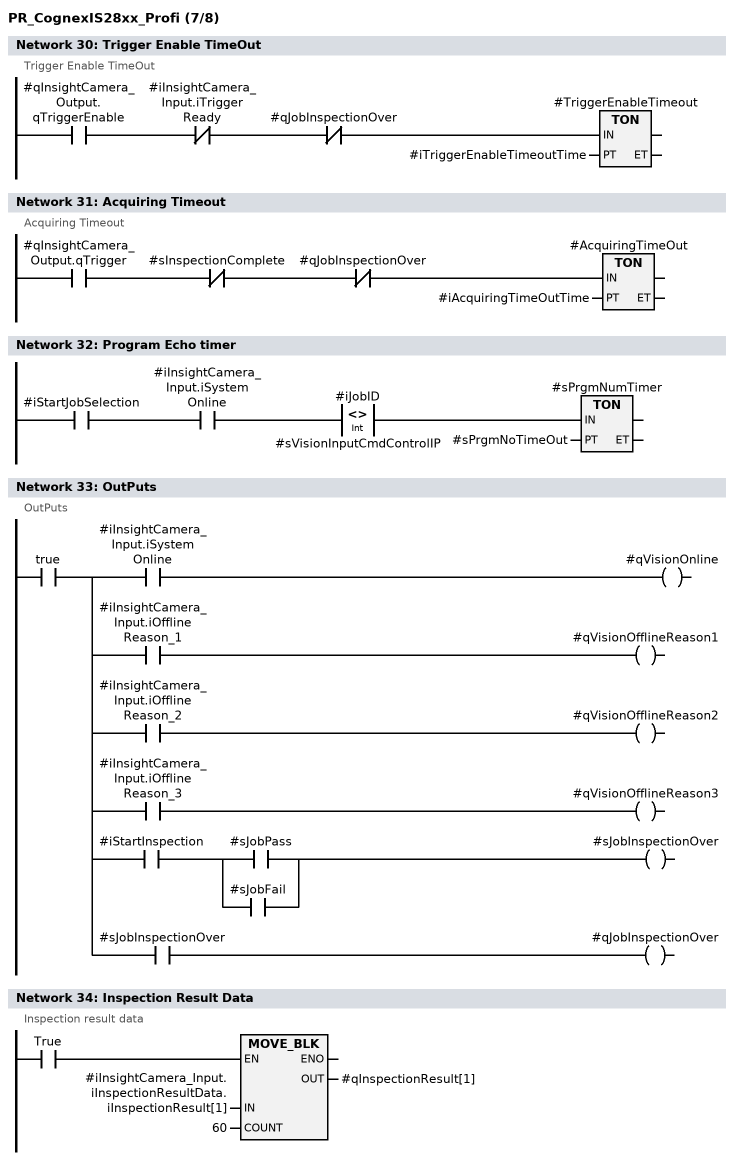
   #TriggerEnableTimeout(IN := #qInsightCamera_Output.qTriggerEnable AND NOT #iInsightCamera_Input.iTriggerReady AND NOT #qJobInspectionOver,   // TON
                         PT := #iTriggerEnableTimeoutTime);
END_REGION

REGION Network 31: Acquiring Timeout
   // Acquiring Timeout
   #AcquiringTimeOut(IN := #qInsightCamera_Output.qTrigger AND NOT #sInspectionComplete AND NOT #qJobInspectionOver,   // TON
                     PT := #iAcquiringTimeOutTime);
END_REGION

REGION Network 32: Program Echo timer
   #sPrgmNumTimer(IN := #iStartJobSelection AND #iInsightCamera_Input.iSystemOnline AND (#iJobID <> #sVisionInputCmdControlIP),   // TON
                  PT := #sPrgmNoTimeOut);
END_REGION

REGION Network 33: OutPuts
   // OutPuts
   RUNG wire#powerrail
      Contact( true )
      wire#w1
      Contact( #iInsightCamera_Input.iSystemOnline )
      Coil( #qVisionOnline )
   END_RUNG
   RUNG wire#w1
      Contact( #iInsightCamera_Input.iOfflineReason_1 )
      Coil( #qVisionOfflineReason1 )
   END_RUNG
   RUNG wire#w1
      Contact( #iInsightCamera_Input.iOfflineReason_2 )
      Coil( #qVisionOfflineReason2 )
   END_RUNG
   RUNG wire#w1
      Contact( #iInsightCamera_Input.iOfflineReason_3 )
      Coil( #qVisionOfflineReason3 )
   END_RUNG
   RUNG wire#w1
      Contact( #iStartInspection )
      wire#w2
      Contact( #sJobPass )
      wire#w3
      Coil( #sJobInspectionOver )
   END_RUNG
   RUNG wire#w2
      Contact( #sJobFail )
   END_RUNG wire#w3
   RUNG wire#w1
      Contact( #sJobInspectionOver )
      Coil( #qJobInspectionOver )
   END_RUNG
   // the same network as SCL:
   #qVisionOnline := true AND #iInsightCamera_Input.iSystemOnline;
   #qVisionOfflineReason1 := true AND #iInsightCamera_Input.iOfflineReason_1;
   #qVisionOfflineReason2 := true AND #iInsightCamera_Input.iOfflineReason_2;
   #qVisionOfflineReason3 := true AND #iInsightCamera_Input.iOfflineReason_3;
   #sJobInspectionOver := true AND #iStartInspection AND (#sJobPass OR #sJobFail);
   #qJobInspectionOver := true AND #sJobInspectionOver;
END_REGION

REGION Network 34: Inspection Result Data
   // Inspection result data
   IF True THEN
       MOVE_BLK(IN := #iInsightCamera_Input.iInspectionResultData.iInspectionResult[1],
                COUNT := 60,
                OUT => #qInspectionResult[1]);
   END_IF;
END_REGION

REGION Network 35: Errors
   // Errors: 
   // qErrTriggerTimeOut: Tigger TimeOut Error Occured
   // qErrAcquiringTimeout: Acquiring TimeOut Error Occured
   // qErrTriggerEnableTimeout: Trigger Enable TimeOut Occured
   // #qErrJobIDEchoMismatch:Job ID Echo Mismatch
   // #qErrJobSelection: Job Error Selection wrong
   // #qErrBothStartOn:Job selection and job inspection both command at time
   // #qErrRetryCount: Retry count value Not set
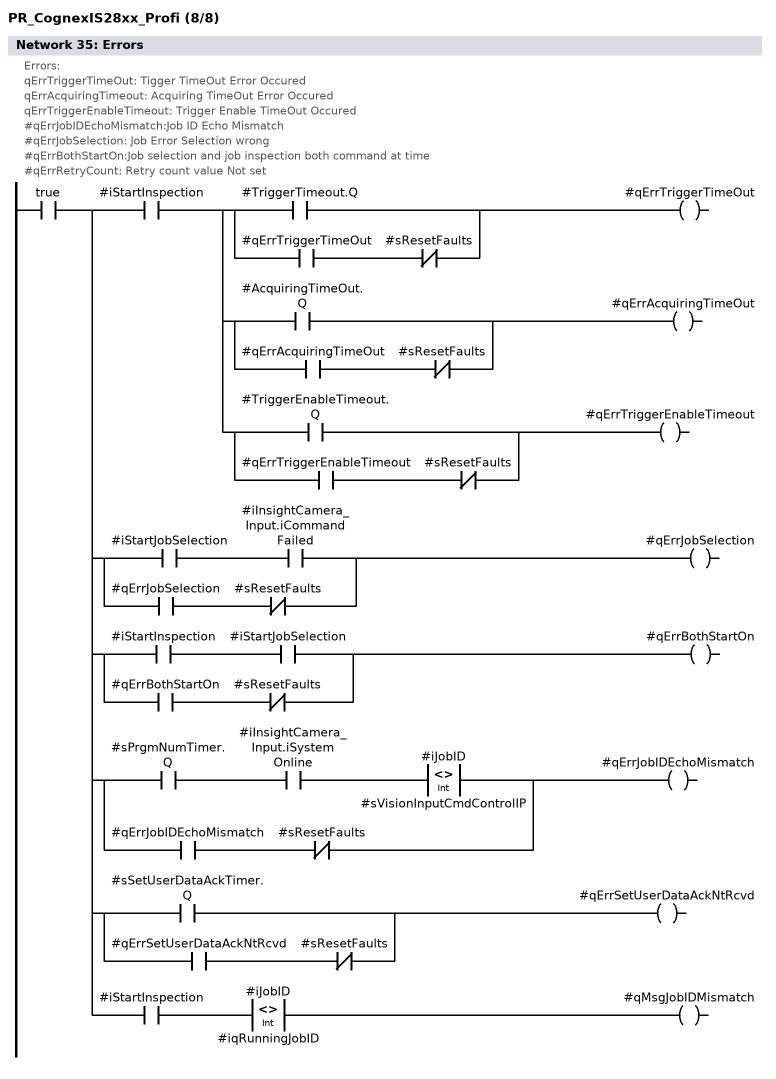
   RUNG wire#powerrail
      Contact( true )
      wire#w1
      Contact( #iStartInspection )
      wire#w2
      Contact( #TriggerTimeout.Q )
      wire#w3
      Coil( #qErrTriggerTimeOut )
   END_RUNG
   RUNG wire#w2
      Contact( #qErrTriggerTimeOut )
      I_Contact( #sResetFaults )
   END_RUNG wire#w3
   RUNG wire#w2
      Contact( #AcquiringTimeOut.Q )
      wire#w4
      Coil( #qErrAcquiringTimeOut )
   END_RUNG
   RUNG wire#w2
      Contact( #qErrAcquiringTimeOut )
      I_Contact( #sResetFaults )
   END_RUNG wire#w4
   RUNG wire#w2
      Contact( #TriggerEnableTimeout.Q )
      wire#w5
      Coil( #qErrTriggerEnableTimeout )
   END_RUNG
   RUNG wire#w2
      Contact( #qErrTriggerEnableTimeout )
      I_Contact( #sResetFaults )
   END_RUNG wire#w5
   RUNG wire#w1
      Contact( #iStartJobSelection )
      Contact( #iInsightCamera_Input.iCommandFailed )
      wire#w6
      Coil( #qErrJobSelection )
   END_RUNG
   RUNG wire#w1
      Contact( #qErrJobSelection )
      I_Contact( #sResetFaults )
   END_RUNG wire#w6
   RUNG wire#w1
      Contact( #iStartInspection )
      Contact( #iStartJobSelection )
      wire#w7
      Coil( #qErrBothStartOn )
   END_RUNG
   RUNG wire#w1
      Contact( #qErrBothStartOn )
      I_Contact( #sResetFaults )
   END_RUNG wire#w7
   RUNG wire#w1
      Contact( #sPrgmNumTimer.Q )
      Contact( #iInsightCamera_Input.iSystemOnline )
      { S7_Templates := "SrcType := Int" } NE_Contact(in1 := #iJobID, in2 := #sVisionInputCmdControlIP)
      wire#w8
      Coil( #qErrJobIDEchoMismatch )
   END_RUNG
   RUNG wire#w1
      Contact( #qErrJobIDEchoMismatch )
      I_Contact( #sResetFaults )
   END_RUNG wire#w8
   RUNG wire#w1
      Contact( #sSetUserDataAckTimer.Q )
      wire#w9
      Coil( #qErrSetUserDataAckNtRcvd )
   END_RUNG
   RUNG wire#w1
      Contact( #qErrSetUserDataAckNtRcvd )
      I_Contact( #sResetFaults )
   END_RUNG wire#w9
   RUNG wire#w1
      Contact( #iStartInspection )
      { S7_Templates := "SrcType := Int" } NE_Contact(in1 := #iJobID, in2 := #iqRunningJobID)
      Coil( #qMsgJobIDMismatch )
   END_RUNG
   // the same network as SCL:
   #_w1 := true AND #iStartInspection;
   #qErrTriggerTimeOut := #_w1 AND (#TriggerTimeout.Q OR (#qErrTriggerTimeOut AND NOT #sResetFaults));
   #qErrAcquiringTimeOut := #_w1 AND (#AcquiringTimeOut.Q OR (#qErrAcquiringTimeOut AND NOT #sResetFaults));
   #qErrTriggerEnableTimeout := #_w1 AND (#TriggerEnableTimeout.Q OR (#qErrTriggerEnableTimeout AND NOT #sResetFaults));
   #qErrJobSelection := true AND ((#iStartJobSelection AND #iInsightCamera_Input.iCommandFailed) OR (#qErrJobSelection AND NOT #sResetFaults));
   #qErrBothStartOn := true AND ((#iStartInspection AND #iStartJobSelection) OR (#qErrBothStartOn AND NOT #sResetFaults));
   #qErrJobIDEchoMismatch := true AND ((#sPrgmNumTimer.Q AND #iInsightCamera_Input.iSystemOnline AND (#iJobID <> #sVisionInputCmdControlIP)) OR (#qErrJobIDEchoMismatch AND NOT #sResetFaults));
   #qErrSetUserDataAckNtRcvd := true AND (#sSetUserDataAckTimer.Q OR (#qErrSetUserDataAckNtRcvd AND NOT #sResetFaults));
   #qMsgJobIDMismatch := true AND #iStartInspection AND (#iJobID <> #iqRunningJobID);
END_REGION
END_FUNCTION_BLOCK

// folder: SM-Modules

FUNCTION "PR_WriteDataSlave" : Void   // FC19, LAD
TITLE = Write Data To Profinet Device
{ S7_Optimized_Access := 'TRUE' }
AUTHOR : GST
FAMILY : SM
NAME : SM0304022002
VERSION : 0.1
   VAR_INPUT
      iNumberOfBytes : Int;   // Number Of Bytes Configured In Hardware
      iSourceStruct : Variant;   // Source Data Structure
   END_VAR
   VAR_OUTPUT
      iOutputAddress : ANY;   // Output Data Address P#Q120.0 BYTE 71
   END_VAR
   VAR_TEMP
      tRetVal : Int;   // Ret Value
      tSrcMovBlck : Array[0..512] of Byte;   // Source Data ARRAY
      tPOS : DInt;   // POS
   END_VAR
BEGIN

REGION Network 1: Header
   // ==============================================================================
   //  Company: Precision Automation & Robotics India Ltd. 
   // ------------------------------------------------------------------------------
   //  Item Code: SM0304022002
   //  Author/Created by: GST
   //  Reviewed/Checked by: Atul P
   //  First Release on: 05-June-2018
   //  Latest update on: 
   // ------------------------------------------------------------------------------
   //  Tested with: CPU firmware, model or simulator testing
   //  Engineering/Editor: TIA Portal V15.1
   // ------------------------------------------------------------------------------
   //  Restrictions: 
   //  Dependencies/Requirements:
   //  This block uses following standard "Siemens" functions:
   // MOVE_BLK_VARIANT
   // Serialize
   // may lead to CPU going to STOP mode.
   // ------------------------------------------------------------------------------
   //  Change Log:
   //  Ver.	Date		Changed by		Details of changes
   //  1.0	05-June-2018	GST                               	First release version
   // ------------------------------------------------------------------------------
   //  Functionality:  This block is used for interface of Write Data From Structure Data To Profinet Device
   // 
   //  Inputs
   // iNumberOfBytes	Int
   // iSourceStruct	Variant
   // 
   //  Outputs
   // iOutputAddress	Any
   // 
   //  In-outs
   //  
   // ------------------------------------------------------------------------------
   //  Errors reported:
   //  1. 
   //  Messages reported:
   //  1. 
   // ==============================================================================
END_REGION

REGION Network 2: Serialize Structure Input Into Array
   // Serialize Structure Input Into Array
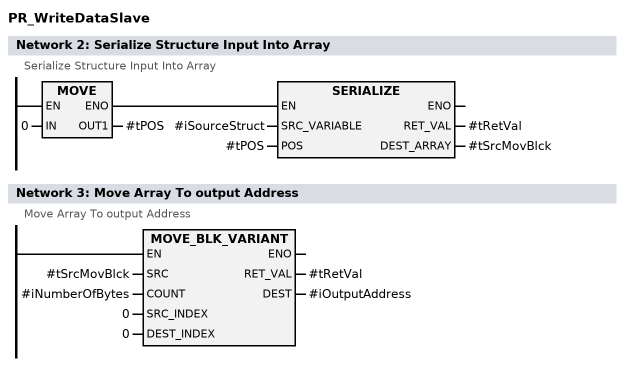
   // no SCL statement known for Serialize: written as a call
   #tPOS := 0;
   #tRetVal := Serialize(SRC_VARIABLE := #iSourceStruct, POS := #tPOS, DEST_ARRAY => #tSrcMovBlck);
END_REGION

REGION Network 3: Move Array To output Address
   // Move Array To output Address
   #tRetVal := MOVE_BLK_VARIANT(SRC := #tSrcMovBlck,
                           COUNT := #iNumberOfBytes,
                           SRC_INDEX := 0,
                           DEST_INDEX := 0,
                           DEST => #iOutputAddress);
END_REGION
END_FUNCTION

FUNCTION "PR_ReadDataSlave" : Void   // FC20, LAD
TITLE = Read Data From Profinet Device
{ S7_Optimized_Access := 'TRUE' }
AUTHOR : GST
FAMILY : SM
NAME : SM0314022001
VERSION : 0.1
// |BLOCK:Cognex Scanner Module
// Item Code : SMxxxxx
// Owner:Precision Automation & Robotics India Ltd.
// Author: GST
// Release Date:05-June-2018
// Version:0.1
// V0.1-Initial release
// |=============================================================================|
// Block Description: This block is used for interface of Read Data From Profinet Device And Store Into Structure DATA
// |=============================================================================|
// Errors:
// 
// =============================================================================|
// Dependency:
// This block uses following standard "Siemens" functions:
// MOVE_BLK_VARIANT
// Deserialize
// may lead to CPU going to STOP mode.
// |
   VAR_INPUT
      iInputAddress : ANY;   // Input Hardware Address P#I120.0 BYTE 77
      iNumberOfBytes : Int;   // Input Number Of Bytes
   END_VAR
   VAR_OUTPUT
      qDestStruct : Variant;   // Destination Data Structure
   END_VAR
   VAR_TEMP
      tRetVal : Int;   // Ret Value
      tDestMovBlck : Array[0..512] of Byte;   // Destination Data Array
      tPOS : DInt;   // POS
   END_VAR
BEGIN

REGION Network 1: Header
   // ==============================================================================
   //  Company: Precision Automation & Robotics India Ltd. 
   // ------------------------------------------------------------------------------
   //  Item Code: SM0314022001
   //  Author/Created by: GST
   //  Reviewed/Checked by: Atul P
   //  First Release on: 05-June-2018
   //  Latest update on:
   // ------------------------------------------------------------------------------
   //  Tested with: CPU firmware, model or simulator testing
   //  Engineering/Editor: TIA Portal V15.1
   // ------------------------------------------------------------------------------
   //  Restrictions: 
   //  Dependencies/Requirements:
   // This block uses following standard "Siemens" functions:
   // MOVE_BLK_VARIANT
   // Deserialize
   // may lead to CPU going to STOP mode.
   // ------------------------------------------------------------------------------
   //  Change Log:
   //  Ver.	Date		Changed by		Details of changes
   //  1.0	05-June-2018	GST                                   	First release version
   // ------------------------------------------------------------------------------
   //  Functionality: This block is used for interface of Read Data From Profinet Device And Store Into Structure DATA
   // 
   //  Inputs
   //  iInputAddress	Any
   // iNumberOfBytes	Int
   // 
   //  Outputs
   // qDestStruct	Variant
   // 
   //  In-outs
   //  
   // ------------------------------------------------------------------------------
   //  Errors reported:
   //  1.
   //  Messages reported:
   //  1. 
   // ==============================================================================
END_REGION

REGION Network 2: Move Input Address Data To Destination Array
   // Move Input Address Data To Destination Array
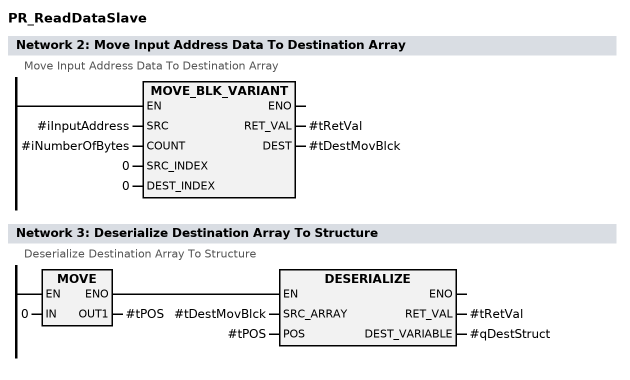
   #tRetVal := MOVE_BLK_VARIANT(SRC := #iInputAddress,
                           COUNT := #iNumberOfBytes,
                           SRC_INDEX := 0,
                           DEST_INDEX := 0,
                           DEST => #tDestMovBlck);
END_REGION

REGION Network 3: Deserialize Destination Array To Structure
   // Deserialize Destination Array To Structure
   // no SCL statement known for Deserialize: written as a call
   #tPOS := 0;
   #tRetVal := Deserialize(SRC_ARRAY := #tDestMovBlck, POS := #tPOS, DEST_VARIABLE => #qDestStruct);
END_REGION
END_FUNCTION